(* IEC 61131-3 sources: plc-st-coding-agent/progress/evidence/f14_v3_parallel_20261112/jobs/custom_deepseek-v4pro (part 2) *)

(* ---- public-hard-05.raw_candidate_02.st ---- *)
FUNCTION_BLOCK MechanicalArmControl
VAR
    Step: INT := 1;                     // Current action step (1..8)
    ActionActive: BOOL := FALSE;        // TRUE when an automated action is being executed
    WaitingForStart: BOOL := TRUE;      // TRUE in single-step mode when waiting for start press
    CycleRunning: BOOL := FALSE;        // TRUE when a cycle is in progress (single/continuous)
    StartPrev: BOOL := FALSE;           // Previous value of Start input for edge detection
    StartPulse: BOOL := FALSE;          // One-scan pulse on rising edge of Start
    WaitingForStartPrev: BOOL := TRUE;  // Snapshot of WaitingForStart at scan start
    CycleRunningPrev: BOOL := FALSE;    // Snapshot of CycleRunning at scan start
END_VAR

// Rising edge detection for Start
StartPulse := Start AND NOT StartPrev;
StartPrev := Start;

// Capture previous states before any logic changes (to avoid race conditions)
WaitingForStartPrev := WaitingForStart;
CycleRunningPrev := CycleRunning;

IF NOT EmergencyStop THEN
    // Emergency stop triggered: stop all actions and reset automated state
    MoveDown := FALSE;
    MoveUp := FALSE;
    MoveLeft := FALSE;
    MoveRight := FALSE;
    ActivateGrip := FALSE;
    ActivateRelease := FALSE;
    Step := 1;
    ActionActive := FALSE;
    WaitingForStart := TRUE;
    CycleRunning := FALSE;
ELSE
    // Normal operation (no emergency stop)
    IF ManualMode THEN
        // Manual mode: direct button control with limit switch interlock
        MoveDown := DownButton AND NOT DownLimitSwitch;
        MoveUp := UpButton AND NOT UpLimitSwitch;
        MoveLeft := LeftButton AND NOT LeftLimitSwitch;
        MoveRight := RightButton AND NOT RightLimitSwitch;
        ActivateGrip := GripButton AND NOT GripLimitSwitch;
        ActivateRelease := ReleaseButton AND NOT ReleaseLimitSwitch;
        // Reset automated state when in manual mode
        Step := 1;
        ActionActive := FALSE;
        WaitingForStart := TRUE;
        CycleRunning := FALSE;
    ELSIF SingleStepMode THEN
        // Single step mode: one action per start press
        MoveDown := FALSE;
        MoveUp := FALSE;
        MoveLeft := FALSE;
        MoveRight := FALSE;
        ActivateGrip := FALSE;
        ActivateRelease := FALSE;

        IF WaitingForStartPrev AND StartPulse THEN
            WaitingForStart := FALSE;
            ActionActive := TRUE;
            Step := 1;  // Always start from step 1
        END_IF;

        IF ActionActive THEN
            CASE Step OF
                1: IF DownLimitSwitch THEN
                       ActionActive := FALSE;
                       WaitingForStart := TRUE;
                       Step := 1;
                   END_IF;
                2: IF GripLimitSwitch THEN
                       ActionActive := FALSE;
                       WaitingForStart := TRUE;
                       Step := 2;
                   END_IF;
                3: IF UpLimitSwitch THEN
                       ActionActive := FALSE;
                       WaitingForStart := TRUE;
                       Step := 3;
                   END_IF;
                4: IF RightLimitSwitch THEN
                       ActionActive := FALSE;
                       WaitingForStart := TRUE;
                       Step := 4;
                   END_IF;
                5: IF DownLimitSwitch THEN
                       ActionActive := FALSE;
                       WaitingForStart := TRUE;
                       Step := 5;
                   END_IF;
                6: IF ReleaseLimitSwitch THEN
                       ActionActive := FALSE;
                       WaitingForStart := TRUE;
                       Step := 6;
                   END_IF;
                7: IF UpLimitSwitch THEN
                       ActionActive := FALSE;
                       WaitingForStart := TRUE;
                       Step := 7;
                   END_IF;
                8: IF LeftLimitSwitch THEN
                       ActionActive := FALSE;
                       WaitingForStart := TRUE;
                       Step := 1;  // Reset to step 1 for next cycle
                   END_IF;
            END_CASE;
        END_IF;

        IF ActionActive THEN
            CASE Step OF
                1: MoveDown := TRUE;
                2: ActivateGrip := TRUE;
                3: MoveUp := TRUE;
                4: MoveRight := TRUE;
                5: MoveDown := TRUE;
                6: ActivateRelease := TRUE;
                7: MoveUp := TRUE;
                8: MoveLeft := TRUE;
            END_CASE;
        END_IF;
    ELSIF SingleCycleMode THEN
        // Single cycle mode: complete one full cycle automatically
        MoveDown := FALSE;
        MoveUp := FALSE;
        MoveLeft := FALSE;
        MoveRight := FALSE;
        ActivateGrip := FALSE;
        ActivateRelease := FALSE;

        IF NOT CycleRunningPrev AND StartPulse THEN
            CycleRunning := TRUE;
            Step := 1;
            ActionActive := TRUE;
        END_IF;

        IF CycleRunning AND ActionActive THEN
            CASE Step OF
                1: IF DownLimitSwitch THEN Step := 2; END_IF;
                2: IF GripLimitSwitch THEN Step := 3; END_IF;
                3: IF UpLimitSwitch THEN Step := 4; END_IF;
                4: IF RightLimitSwitch THEN Step := 5; END_IF;
                5: IF DownLimitSwitch THEN Step := 6; END_IF;
                6: IF ReleaseLimitSwitch THEN Step := 7; END_IF;
                7: IF UpLimitSwitch THEN Step := 8; END_IF;
                8: IF LeftLimitSwitch THEN
                       ActionActive := FALSE;   // Cycle finished
                       CycleRunning := FALSE;
                       Step := 1;               // Reset for next start
                   END_IF;
            END_CASE;
        END_IF;

        IF CycleRunning AND ActionActive THEN
            CASE Step OF
                1: MoveDown := TRUE;
                2: ActivateGrip := TRUE;
                3: MoveUp := TRUE;
                4: MoveRight := TRUE;
                5: MoveDown := TRUE;
                6: ActivateRelease := TRUE;
                7: MoveUp := TRUE;
                8: MoveLeft := TRUE;
            END_CASE;
        END_IF;
    ELSIF ContinuousMode THEN
        // Continuous mode: repeat cycle indefinitely
        MoveDown := FALSE;
        MoveUp := FALSE;
        MoveLeft := FALSE;
        MoveRight := FALSE;
        ActivateGrip := FALSE;
        ActivateRelease := FALSE;

        IF NOT CycleRunningPrev AND StartPulse THEN
            CycleRunning := TRUE;
            Step := 1;
            ActionActive := TRUE;
        END_IF;

        IF CycleRunning AND ActionActive THEN
            CASE Step OF
                1: IF DownLimitSwitch THEN Step := 2; END_IF;
                2: IF GripLimitSwitch THEN Step := 3; END_IF;
                3: IF UpLimitSwitch THEN Step := 4; END_IF;
                4: IF RightLimitSwitch THEN Step := 5; END_IF;
                5: IF DownLimitSwitch THEN Step := 6; END_IF;
                6: IF ReleaseLimitSwitch THEN Step := 7; END_IF;
                7: IF UpLimitSwitch THEN Step := 8; END_IF;
                8: IF LeftLimitSwitch THEN Step := 1; END_IF;  // Loop back
            END_CASE;
        END_IF;

        IF CycleRunning AND ActionActive THEN
            CASE Step OF
                1: MoveDown := TRUE;
                2: ActivateGrip := TRUE;
                3: MoveUp := TRUE;
                4: MoveRight := TRUE;
                5: MoveDown := TRUE;
                6: ActivateRelease := TRUE;
                7: MoveUp := TRUE;
                8: MoveLeft := TRUE;
            END_CASE;
        END_IF;
    ELSE
        // No mode selected (should not happen, but safe default)
        MoveDown := FALSE;
        MoveUp := FALSE;
        MoveLeft := FALSE;
        MoveRight := FALSE;
        ActivateGrip := FALSE;
        ActivateRelease := FALSE;
        Step := 1;
        ActionActive := FALSE;
        WaitingForStart := TRUE;
        CycleRunning := FALSE;
    END_IF;
END_IF;

END_FUNCTION_BLOCK

(* ---- public-hard-06.candidate_01.st ---- *)
TYPE T_PRODUCTION_STATE :
(
    IDLE,
    MOVING_FEED_TO_WASH,
    AT_WASH,
    MOVING_WASH_TO_WEIGHT,
    AT_WEIGHT_WAIT,
    AT_WEIGHT_REJECT,
    MOVING_WEIGHT_TO_FIRING,
    AT_FIRING,
    MOVING_FIRING_TO_OUTPUT,
    AT_OUTPUT
);
END_TYPE;

FUNCTION_BLOCK ProductionControl
VAR_INPUT
    Mode : BOOL;
    ForwardButton : BOOL;
    ReverseButton : BOOL;
    SensorFeed : BOOL;
    SensorWash : BOOL;
    SensorWeight : BOOL;
    SensorFiring : BOOL;
    SensorOutput : BOOL;
    washComplete : BOOL;
    weightComplete : BOOL;
    weight : REAL;
    firingComplete : BOOL;
END_VAR
VAR_OUTPUT
    MotorForward : BOOL;
    MotorReverse : BOOL;
    kick : BOOL;
    CompletionLight : BOOL;
    firingTemp : REAL;
END_VAR
VAR
    currentState : T_PRODUCTION_STATE := IDLE;
END_VAR

(* ---- public-hard-06.candidate_02.st ---- *)
TYPE T_PRODUCTION_STATE :
(
    IDLE,
    MOVING_FEED_TO_WASH,
    AT_WASH,
    MOVING_WASH_TO_WEIGHT,
    AT_WEIGHT_WAIT,
    AT_WEIGHT_REJECT,
    MOVING_WEIGHT_TO_FIRING,
    AT_FIRING,
    MOVING_FIRING_TO_OUTPUT,
    AT_OUTPUT
);
END_TYPE;

FUNCTION_BLOCK ProductionControl
VAR_INPUT
    Mode : BOOL;
    ForwardButton : BOOL;
    ReverseButton : BOOL;
    SensorFeed : BOOL;
    SensorWash : BOOL;
    SensorWeight : BOOL;
    SensorFiring : BOOL;
    SensorOutput : BOOL;
    washComplete : BOOL;
    weightComplete : BOOL;
    weight : REAL;
    firingComplete : BOOL;
END_VAR
VAR_OUTPUT
    MotorForward : BOOL;
    MotorReverse : BOOL;
    kick : BOOL;
    CompletionLight : BOOL;
    firingTemp : REAL;
END_VAR
VAR
    currentState : T_PRODUCTION_STATE := IDLE;
END_VAR

IF Mode = FALSE THEN
    // Manual mode
    IF ForwardButton AND NOT ReverseButton THEN
        MotorForward := TRUE;
        MotorReverse := FALSE;
    ELSIF ReverseButton AND NOT ForwardButton THEN
        MotorForward := FALSE;
        MotorReverse := TRUE;
    ELSE
        MotorForward := FALSE;
        MotorReverse := FALSE;
    END_IF;
    // Reset all automatic outputs and state
    kick := FALSE;
    CompletionLight := FALSE;
    firingTemp := 0.0;
    currentState := IDLE;
ELSE
    // Automatic mode
    // Set default outputs for this scan
    MotorReverse := FALSE;
    MotorForward := FALSE;
    kick := FALSE;
    CompletionLight := FALSE;
    // firingTemp retains its last calculated value unless updated in qualified weighing

    CASE currentState OF
        IDLE:
            IF SensorFeed THEN
                currentState := MOVING_FEED_TO_WASH;
                MotorForward := TRUE;
            END_IF;

        MOVING_FEED_TO_WASH:
            MotorForward := TRUE;
            IF SensorWash THEN
                MotorForward := FALSE;
                currentState := AT_WASH;
            END_IF;

        AT_WASH:
            IF washComplete THEN
                MotorForward := TRUE;
                currentState := MOVING_WASH_TO_WEIGHT;
            END_IF;

        MOVING_WASH_TO_WEIGHT:
            MotorForward := TRUE;
            IF SensorWeight THEN
                MotorForward := FALSE;
                currentState := AT_WEIGHT_WAIT;
            END_IF;

        AT_WEIGHT_WAIT:
            IF weightComplete THEN
                IF (weight >= 100.0) AND (weight <= 200.0) THEN
                    // Qualified material
                    firingTemp := 500.0 + (weight - 100.0) * 0.5;
                    MotorForward := TRUE;
                    currentState := MOVING_WEIGHT_TO_FIRING;
                ELSE
                    // Unqualified material
                    kick := TRUE;
                    currentState := AT_WEIGHT_REJECT;
                END_IF;
            END_IF;

        AT_WEIGHT_REJECT:
            kick := TRUE;
            IF NOT SensorWeight THEN
                kick := FALSE;
                currentState := IDLE;
            END_IF;

        MOVING_WEIGHT_TO_FIRING:
            MotorForward := TRUE;
            IF SensorFiring THEN
                MotorForward := FALSE;
                currentState := AT_FIRING;
            END_IF;

        AT_FIRING:
            IF firingComplete THEN
                MotorForward := TRUE;
                currentState := MOVING_FIRING_TO_OUTPUT;
            END_IF;

        MOVING_FIRING_TO_OUTPUT:
            MotorForward := TRUE;
            IF SensorOutput THEN
                MotorForward := FALSE;
                currentState := AT_OUTPUT;
            END_IF;

        AT_OUTPUT:
            CompletionLight := TRUE;
            IF NOT SensorOutput THEN
                CompletionLight := FALSE;
                currentState := IDLE;
            END_IF;
    END_CASE;
END_IF;

END_FUNCTION_BLOCK

(* ---- public-hard-06.raw_candidate_01.st ---- *)
TYPE T_PRODUCTION_STATE :
(
    IDLE,
    MOVING_FEED_TO_WASH,
    AT_WASH,
    MOVING_WASH_TO_WEIGHT,
    AT_WEIGHT_WAIT,
    AT_WEIGHT_REJECT,
    MOVING_WEIGHT_TO_FIRING,
    AT_FIRING,
    MOVING_FIRING_TO_OUTPUT,
    AT_OUTPUT
);
END_TYPE

FUNCTION_BLOCK ProductionControl
VAR_INPUT
    Mode : BOOL;
    ForwardButton : BOOL;
    ReverseButton : BOOL;
    SensorFeed : BOOL;
    SensorWash : BOOL;
    SensorWeight : BOOL;
    SensorFiring : BOOL;
    SensorOutput : BOOL;
    washComplete : BOOL;
    weightComplete : BOOL;
    weight : REAL;
    firingComplete : BOOL;
END_VAR
VAR_OUTPUT
    MotorForward : BOOL;
    MotorReverse : BOOL;
    kick : BOOL;
    CompletionLight : BOOL;
    firingTemp : REAL;
END_VAR
VAR
    currentState : T_PRODUCTION_STATE := IDLE;
END_VAR

(* ---- public-hard-06.raw_candidate_02.st ---- *)
TYPE T_PRODUCTION_STATE :
(
    IDLE,
    MOVING_FEED_TO_WASH,
    AT_WASH,
    MOVING_WASH_TO_WEIGHT,
    AT_WEIGHT_WAIT,
    AT_WEIGHT_REJECT,
    MOVING_WEIGHT_TO_FIRING,
    AT_FIRING,
    MOVING_FIRING_TO_OUTPUT,
    AT_OUTPUT
);
END_TYPE;

FUNCTION_BLOCK ProductionControl
VAR_INPUT
    Mode : BOOL;
    ForwardButton : BOOL;
    ReverseButton : BOOL;
    SensorFeed : BOOL;
    SensorWash : BOOL;
    SensorWeight : BOOL;
    SensorFiring : BOOL;
    SensorOutput : BOOL;
    washComplete : BOOL;
    weightComplete : BOOL;
    weight : REAL;
    firingComplete : BOOL;
END_VAR
VAR_OUTPUT
    MotorForward : BOOL;
    MotorReverse : BOOL;
    kick : BOOL;
    CompletionLight : BOOL;
    firingTemp : REAL;
END_VAR
VAR
    currentState : T_PRODUCTION_STATE := IDLE;
END_VAR

IF Mode = FALSE THEN
    // Manual mode
    IF ForwardButton AND NOT ReverseButton THEN
        MotorForward := TRUE;
        MotorReverse := FALSE;
    ELSIF ReverseButton AND NOT ForwardButton THEN
        MotorForward := FALSE;
        MotorReverse := TRUE;
    ELSE
        MotorForward := FALSE;
        MotorReverse := FALSE;
    END_IF;
    // Reset all automatic outputs and state
    kick := FALSE;
    CompletionLight := FALSE;
    firingTemp := 0.0;
    currentState := IDLE;
ELSE
    // Automatic mode
    // Set default outputs for this scan
    MotorReverse := FALSE;
    MotorForward := FALSE;
    kick := FALSE;
    CompletionLight := FALSE;
    // firingTemp retains its last calculated value unless updated in qualified weighing

    CASE currentState OF
        IDLE:
            IF SensorFeed THEN
                currentState := MOVING_FEED_TO_WASH;
                MotorForward := TRUE;
            END_IF;

        MOVING_FEED_TO_WASH:
            MotorForward := TRUE;
            IF SensorWash THEN
                MotorForward := FALSE;
                currentState := AT_WASH;
            END_IF;

        AT_WASH:
            IF washComplete THEN
                MotorForward := TRUE;
                currentState := MOVING_WASH_TO_WEIGHT;
            END_IF;

        MOVING_WASH_TO_WEIGHT:
            MotorForward := TRUE;
            IF SensorWeight THEN
                MotorForward := FALSE;
                currentState := AT_WEIGHT_WAIT;
            END_IF;

        AT_WEIGHT_WAIT:
            IF weightComplete THEN
                IF (weight >= 100.0) AND (weight <= 200.0) THEN
                    // Qualified material
                    firingTemp := 500.0 + (weight - 100.0) * 0.5;
                    MotorForward := TRUE;
                    currentState := MOVING_WEIGHT_TO_FIRING;
                ELSE
                    // Unqualified material
                    kick := TRUE;
                    currentState := AT_WEIGHT_REJECT;
                END_IF;
            END_IF;

        AT_WEIGHT_REJECT:
            kick := TRUE;
            IF NOT SensorWeight THEN
                kick := FALSE;
                currentState := IDLE;
            END_IF;

        MOVING_WEIGHT_TO_FIRING:
            MotorForward := TRUE;
            IF SensorFiring THEN
                MotorForward := FALSE;
                currentState := AT_FIRING;
            END_IF;

        AT_FIRING:
            IF firingComplete THEN
                MotorForward := TRUE;
                currentState := MOVING_FIRING_TO_OUTPUT;
            END_IF;

        MOVING_FIRING_TO_OUTPUT:
            MotorForward := TRUE;
            IF SensorOutput THEN
                MotorForward := FALSE;
                currentState := AT_OUTPUT;
            END_IF;

        AT_OUTPUT:
            CompletionLight := TRUE;
            IF NOT SensorOutput THEN
                CompletionLight := FALSE;
                currentState := IDLE;
            END_IF;
    END_CASE;
END_IF;

END_FUNCTION_BLOCK

(* ---- public-medium-01.candidate_01.st ---- *)
TYPE ST_Pump :
STRUCT
    priority : INT;
    selection : BOOL;
    RunComd : BOOL;
END_STRUCT;
END_TYPE;

FUNCTION_BLOCK FB_MultiPumpControl
VAR_INPUT
    mode : BOOL;
    start : BOOL;
    stop : BOOL;
END_VAR
VAR_IN_OUT
    pumpGroup : ARRAY[1..5] OF ST_Pump;
END_VAR
VAR
    runActive : BOOL := FALSE;
    autoSelected : ARRAY[1..5] OF BOOL;
    i : INT;
    j : INT;
    rank : INT;
END_VAR

IF stop THEN
    runActive := FALSE;
    FOR i := 1 TO 5 DO
        pumpGroup[i].RunComd := FALSE;
    END_FOR;
ELSE
    IF start THEN
        runActive := TRUE;
    END_IF;

    IF runActive THEN
        IF mode THEN
            FOR i := 1 TO 5 DO
                rank := 0;
                FOR j := 1 TO 5 DO
                    IF (pumpGroup[j].priority > pumpGroup[i].priority) OR
                       ((pumpGroup[j].priority = pumpGroup[i].priority) AND (j < i)) THEN
                        rank := rank + 1;
                    END_IF;
                END_FOR;
                autoSelected[i] := (rank < 3);
            END_FOR;

            FOR i := 1 TO 5 DO
                pumpGroup[i].RunComd := autoSelected[i];
            END_FOR;
        ELSE
            FOR i := 1 TO 5 DO
                pumpGroup[i].RunComd := pumpGroup[i].selection;
            END_FOR;
        END_IF;
    ELSE
        FOR i := 1 TO 5 DO
            pumpGroup[i].RunComd := FALSE;
        END_FOR;
    END_IF;
END_IF;

END_FUNCTION_BLOCK

(* ---- public-medium-01.candidate_02.st ---- *)
TYPE ST_Pump :
STRUCT
    priority : INT;
    selection : BOOL;
    RunComd : BOOL;
END_STRUCT;
END_TYPE;

FUNCTION_BLOCK FB_MultiPumpControl
VAR_INPUT
    mode : BOOL;
    start : BOOL;
    stop : BOOL;
END_VAR
VAR_IN_OUT
    pumpGroup : ARRAY[1..5] OF ST_Pump;
END_VAR
VAR
    runActive : BOOL := FALSE;
    autoSelected : ARRAY[1..5] OF BOOL;
    i : INT;
    j : INT;
    rank : INT;
END_VAR

IF stop THEN
    runActive := FALSE;
    FOR i := 1 TO 5 DO
        pumpGroup[i].RunComd := FALSE;
    END_FOR;
ELSE
    IF start THEN
        runActive := TRUE;
    END_IF;

    IF runActive THEN
        IF mode THEN
            FOR i := 1 TO 5 DO
                rank := 0;
                FOR j := 1 TO 5 DO
                    IF (pumpGroup[j].priority > pumpGroup[i].priority) OR
                       ((pumpGroup[j].priority = pumpGroup[i].priority) AND (j < i)) THEN
                        rank := rank + 1;
                    END_IF;
                END_FOR;
                autoSelected[i] := (rank < 3);
            END_FOR;

            FOR i := 1 TO 5 DO
                pumpGroup[i].RunComd := autoSelected[i];
            END_FOR;
        ELSE
            FOR i := 1 TO 5 DO
                pumpGroup[i].RunComd := pumpGroup[i].selection;
            END_FOR;
        END_IF;
    ELSE
        FOR i := 1 TO 5 DO
            pumpGroup[i].RunComd := FALSE;
        END_FOR;
    END_IF;
END_IF;

END_FUNCTION_BLOCK

(* ---- public-medium-01.raw_candidate_01.st ---- *)
TYPE ST_Pump :
STRUCT
    priority : INT;
    selection : BOOL;
    RunComd : BOOL;
END_STRUCT;
END_TYPE;

FUNCTION_BLOCK FB_MultiPumpControl
VAR_INPUT
    mode : BOOL;
    start : BOOL;
    stop : BOOL;
END_VAR
VAR_IN_OUT
    pumpGroup : ARRAY[1..5] OF ST_Pump;
END_VAR
VAR
    runActive : BOOL := FALSE;
    autoSelected : ARRAY[1..5] OF BOOL;
    i : INT;
    j : INT;
    rank : INT;
END_VAR

IF stop THEN
    runActive := FALSE;
    FOR i := 1 TO 5 DO
        pumpGroup[i].RunComd := FALSE;
    END_FOR;
ELSE
    IF start THEN
        runActive := TRUE;
    END_IF;

    IF runActive THEN
        IF mode THEN
            FOR i := 1 TO 5 DO
                rank := 0;
                FOR j := 1 TO 5 DO
                    IF (pumpGroup[j].priority > pumpGroup[i].priority) OR
                       ((pumpGroup[j].priority = pumpGroup[i].priority) AND (j < i)) THEN
                        rank := rank + 1;
                    END_IF;
                END_FOR;
                autoSelected[i] := (rank < 3);
            END_FOR;

            FOR i := 1 TO 5 DO
                pumpGroup[i].RunComd := autoSelected[i];
            END_FOR;
        ELSE
            FOR i := 1 TO 5 DO
                pumpGroup[i].RunComd := pumpGroup[i].selection;
            END_FOR;
        END_IF;
    ELSE
        FOR i := 1 TO 5 DO
            pumpGroup[i].RunComd := FALSE;
        END_FOR;
    END_IF;
END_IF;

END_FUNCTION_BLOCK

(* ---- public-medium-01.raw_candidate_02.st ---- *)
TYPE ST_Pump :
STRUCT
    priority : INT;
    selection : BOOL;
    RunComd : BOOL;
END_STRUCT
END_TYPE

FUNCTION_BLOCK FB_MultiPumpControl
VAR_INPUT
    mode : BOOL;
    start : BOOL;
    stop : BOOL;
END_VAR
VAR_IN_OUT
    pumpGroup : ARRAY[1..5] OF ST_Pump;
END_VAR
VAR
    runActive : BOOL := FALSE;
    autoSelected : ARRAY[1..5] OF BOOL;
    i : INT;
    j : INT;
    rank : INT;
END_VAR

IF stop THEN
    runActive := FALSE;
    FOR i := 1 TO 5 DO
        pumpGroup[i].RunComd := FALSE;
    END_FOR;
ELSE
    IF start THEN
        runActive := TRUE;
    END_IF;

    IF runActive THEN
        IF mode THEN
            FOR i := 1 TO 5 DO
                rank := 0;
                FOR j := 1 TO 5 DO
                    IF (pumpGroup[j].priority > pumpGroup[i].priority) OR
                       ((pumpGroup[j].priority = pumpGroup[i].priority) AND (j < i)) THEN
                        rank := rank + 1;
                    END_IF;
                END_FOR;
                autoSelected[i] := (rank < 3);
            END_FOR;

            FOR i := 1 TO 5 DO
                pumpGroup[i].RunComd := autoSelected[i];
            END_FOR;
        ELSE
            FOR i := 1 TO 5 DO
                pumpGroup[i].RunComd := pumpGroup[i].selection;
            END_FOR;
        END_IF;
    ELSE
        FOR i := 1 TO 5 DO
            pumpGroup[i].RunComd := FALSE;
        END_FOR;
    END_IF;
END_IF;

END_FUNCTION_BLOCK

(* ---- public-medium-02.candidate_01.st ---- *)
TYPE ST_AnalogChannel :
STRUCT
    enable : BOOL;
    hiLIM : REAL;
    loLIM : REAL;
    bipolar : BOOL;
    measuringMode : INT;
    retVal : WORD;
    outputValue : REAL;
END_STRUCT;
END_TYPE;

FUNCTION_BLOCK AnalogBatchProcessing
VAR_INPUT
    count : DINT;
END_VAR
VAR_INOUT
    analogValues : ARRAY[*] OF INT;
    channels : ARRAY[*] OF ST_AnalogChannel;
END_VAR
VAR
    i : DINT;
    idxA : DINT;
    idxC : DINT;
    lbA : DINT;
    lbC : DINT;
    raw : INT;
    rawReal : REAL;
    rawMin : REAL;
    rawSpan : REAL;
    engSpan : REAL;
END_VAR

    lbA := LOWER_BOUND(analogValues, 1);
    lbC := LOWER_BOUND(channels, 1);

    FOR i := 0 TO count - 1 DO
        idxA := lbA + i;
        idxC := lbC + i;
        raw := analogValues[idxA];
        channels[idxC].retVal := 0;

        IF channels[idxC].enable THEN
            IF channels[idxC].measuringMode <> 0 AND channels[idxC].measuringMode <> 1 AND channels[idxC].measuringMode <> 2 THEN
                channels[idxC].retVal := WORD#16#8001;
            ELSIF channels[idxC].hiLIM <= channels[idxC].loLIM THEN
                channels[idxC].retVal := WORD#16#8002;
            ELSIF channels[idxC].measuringMode = 0 THEN
                rawReal := INT_TO_REAL(raw);

                IF channels[idxC].bipolar THEN
                    rawMin := -27648.0;
                    rawSpan := 55296.0;
                ELSE
                    rawMin := 0.0;
                    rawSpan := 27648.0;
                END_IF;

                engSpan := channels[idxC].hiLIM - channels[idxC].loLIM;
                channels[idxC].outputValue := channels[idxC].loLIM + (rawReal - rawMin) * engSpan / rawSpan;
            ELSIF channels[idxC].measuringMode = 1 THEN
                rawReal := INT_TO_REAL(raw);
                channels[idxC].outputValue := rawReal / 10.0;
            ELSE
                rawReal := INT_TO_REAL(raw);
                channels[idxC].outputValue := rawReal / 100.0;
            END_IF;
        END_IF;
    END_FOR;

END_FUNCTION_BLOCK

(* ---- public-medium-02.candidate_02.st ---- *)
TYPE ST_AnalogChannel :
STRUCT
    enable : BOOL;
    hiLIM : REAL;
    loLIM : REAL;
    bipolar : BOOL;
    measuringMode : INT;
    retVal : WORD;
    outputValue : REAL;
END_STRUCT;
END_TYPE;

FUNCTION_BLOCK AnalogBatchProcessing
VAR_INPUT
    count : DINT;
END_VAR
VAR_IN_OUT
    analogValues : ARRAY[*] OF INT;
    channels : ARRAY[*] OF ST_AnalogChannel;
END_VAR
VAR
    i : DINT;
    idxA : DINT;
    idxC : DINT;
    lbA : DINT;
    lbC : DINT;
    raw : INT;
    rawReal : REAL;
    rawMin : REAL;
    rawSpan : REAL;
    engSpan : REAL;
END_VAR

    lbA := LOWER_BOUND(analogValues, 1);
    lbC := LOWER_BOUND(channels, 1);

    FOR i := 0 TO count - 1 DO
        idxA := lbA + i;
        idxC := lbC + i;

        IF channels[idxC].enable THEN
            IF channels[idxC].measuringMode <> 0 AND channels[idxC].measuringMode <> 1 AND channels[idxC].measuringMode <> 2 THEN
                channels[idxC].retVal := WORD#16#8001;
            ELSIF channels[idxC].hiLIM <= channels[idxC].loLIM THEN
                channels[idxC].retVal := WORD#16#8002;
            ELSE
                raw := analogValues[idxA];
                rawReal := INT_TO_REAL(raw);
                CASE channels[idxC].measuringMode OF
                    0:
                        IF channels[idxC].bipolar THEN
                            rawMin := -27648.0;
                            rawSpan := 55296.0;
                        ELSE
                            rawMin := 0.0;
                            rawSpan := 27648.0;
                        END_IF;
                        engSpan := channels[idxC].hiLIM - channels[idxC].loLIM;
                        channels[idxC].outputValue := channels[idxC].loLIM + (rawReal - rawMin) * engSpan / rawSpan;
                    1:
                        channels[idxC].outputValue := rawReal / 10.0;
                    2:
                        channels[idxC].outputValue := rawReal / 100.0;
                END_CASE;
                channels[idxC].retVal := 0;
            END_IF;
        END_IF;
    END_FOR;

END_FUNCTION_BLOCK

(* ---- public-medium-02.raw_candidate_01.st ---- *)
TYPE ST_AnalogChannel :
STRUCT
    enable : BOOL;
    hiLIM : REAL;
    loLIM : REAL;
    bipolar : BOOL;
    measuringMode : INT;
    retVal : WORD;
    outputValue : REAL;
END_STRUCT
END_TYPE

FUNCTION_BLOCK AnalogBatchProcessing
VAR_INPUT
    count : DINT;
END_VAR
VAR_INOUT
    analogValues : ARRAY[*] OF INT;
    channels : ARRAY[*] OF ST_AnalogChannel;
END_VAR
VAR
    i : DINT;
    idxA : DINT;
    idxC : DINT;
    lbA : DINT;
    lbC : DINT;
    raw : INT;
    rawReal : REAL;
    rawMin : REAL;
    rawSpan : REAL;
    engSpan : REAL;
END_VAR

    lbA := LOWER_BOUND(analogValues, 1);
    lbC := LOWER_BOUND(channels, 1);

    FOR i := 0 TO count - 1 DO
        idxA := lbA + i;
        idxC := lbC + i;
        raw := analogValues[idxA];
        channels[idxC].retVal := 0;

        IF channels[idxC].enable THEN
            IF channels[idxC].measuringMode <> 0 AND channels[idxC].measuringMode <> 1 AND channels[idxC].measuringMode <> 2 THEN
                channels[idxC].retVal := WORD#16#8001;
            ELSIF channels[idxC].hiLIM <= channels[idxC].loLIM THEN
                channels[idxC].retVal := WORD#16#8002;
            ELSIF channels[idxC].measuringMode = 0 THEN
                rawReal := INT_TO_REAL(raw);

                IF channels[idxC].bipolar THEN
                    rawMin := -27648.0;
                    rawSpan := 55296.0;
                ELSE
                    rawMin := 0.0;
                    rawSpan := 27648.0;
                END_IF

                engSpan := channels[idxC].hiLIM - channels[idxC].loLIM;
                channels[idxC].outputValue := channels[idxC].loLIM + (rawReal - rawMin) * engSpan / rawSpan;
            ELSIF channels[idxC].measuringMode = 1 THEN
                rawReal := INT_TO_REAL(raw);
                channels[idxC].outputValue := rawReal / 10.0;
            ELSE
                rawReal := INT_TO_REAL(raw);
                channels[idxC].outputValue := rawReal / 100.0;
            END_IF
        END_IF
    END_FOR

END_FUNCTION_BLOCK

(* ---- public-medium-02.raw_candidate_02.st ---- *)
TYPE ST_AnalogChannel :
STRUCT
    enable : BOOL;
    hiLIM : REAL;
    loLIM : REAL;
    bipolar : BOOL;
    measuringMode : INT;
    retVal : WORD;
    outputValue : REAL;
END_STRUCT;
END_TYPE;

FUNCTION_BLOCK AnalogBatchProcessing
VAR_INPUT
    count : DINT;
END_VAR
VAR_IN_OUT
    analogValues : ARRAY[*] OF INT;
    channels : ARRAY[*] OF ST_AnalogChannel;
END_VAR
VAR
    i : DINT;
    idxA : DINT;
    idxC : DINT;
    lbA : DINT;
    lbC : DINT;
    raw : INT;
    rawReal : REAL;
    rawMin : REAL;
    rawSpan : REAL;
    engSpan : REAL;
END_VAR

    lbA := LOWER_BOUND(analogValues, 1);
    lbC := LOWER_BOUND(channels, 1);

    FOR i := 0 TO count - 1 DO
        idxA := lbA + i;
        idxC := lbC + i;

        IF channels[idxC].enable THEN
            IF channels[idxC].measuringMode <> 0 AND channels[idxC].measuringMode <> 1 AND channels[idxC].measuringMode <> 2 THEN
                channels[idxC].retVal := WORD#16#8001;
            ELSIF channels[idxC].hiLIM <= channels[idxC].loLIM THEN
                channels[idxC].retVal := WORD#16#8002;
            ELSE
                raw := analogValues[idxA];
                rawReal := INT_TO_REAL(raw);
                CASE channels[idxC].measuringMode OF
                    0:
                        IF channels[idxC].bipolar THEN
                            rawMin := -27648.0;
                            rawSpan := 55296.0;
                        ELSE
                            rawMin := 0.0;
                            rawSpan := 27648.0;
                        END_IF;
                        engSpan := channels[idxC].hiLIM - channels[idxC].loLIM;
                        channels[idxC].outputValue := channels[idxC].loLIM + (rawReal - rawMin) * engSpan / rawSpan;
                    1:
                        channels[idxC].outputValue := rawReal / 10.0;
                    2:
                        channels[idxC].outputValue := rawReal / 100.0;
                END_CASE;
                channels[idxC].retVal := 0;
            END_IF;
        END_IF;
    END_FOR;

END_FUNCTION_BLOCK

(* ---- public-medium-03.candidate_01.st ---- *)
FUNCTION_BLOCK FB_MovingAverage
VAR_INPUT
    cyclicExecution : BOOL;
    trigger : BOOL;
    value : LREAL;
    windowSize : INT;
    reset : BOOL;
END_VAR
VAR_OUTPUT
    average : LREAL;
    windowSizeReached : BOOL;
    error : BOOL;
    status : WORD;
END_VAR
VAR
    buffer : ARRAY[0..99] OF LREAL;
    count : INT := 0;
    writeIndex : INT := 0;
    sum : LREAL := 0.0;
    prevTrigger : BOOL := FALSE;
    prevWindowSize : INT := 0;
    updateNow : BOOL;
END_VAR

IF (windowSize < 1) OR (windowSize > 100) THEN
    error := TRUE;
    status := 16#8200;
    average := 0.0;
    windowSizeReached := FALSE;
    count := 0;
    writeIndex := 0;
    sum := 0.0;
ELSE
    error := FALSE;
    status := 16#0000;

    IF reset OR (windowSize <> prevWindowSize) THEN
        count := 0;
        writeIndex := 0;
        sum := 0.0;
        average := 0.0;
        windowSizeReached := FALSE;
    END_IF;
    prevWindowSize := windowSize;

    IF cyclicExecution THEN
        updateNow := TRUE;
    ELSIF (trigger AND NOT prevTrigger) THEN
        updateNow := TRUE;
    ELSE
        updateNow := FALSE;
    END_IF;

    IF updateNow THEN
        IF count < windowSize THEN
            buffer[writeIndex] := value;
            sum := sum + value;
            count := count + 1;
            writeIndex := writeIndex + 1;
        ELSE
            sum := sum - buffer[writeIndex] + value;
            buffer[writeIndex] := value;
            writeIndex := (writeIndex + 1) MOD windowSize;
        END_IF;
        IF count > 0 THEN
            average := sum / count;
        ELSE
            average := 0.0;
        END_IF;
        windowSizeReached := (count >= windowSize);
    END_IF;
END_IF;

prevTrigger := trigger;

(* ---- public-medium-03.candidate_02.st ---- *)
FUNCTION_BLOCK FB_MovingAverage
VAR_INPUT
    cyclicExecution : BOOL;
    trigger : BOOL;
    value : LREAL;
    windowSize : INT;
    reset : BOOL;
END_VAR
VAR_OUTPUT
    average : LREAL;
    windowSizeReached : BOOL;
    error : BOOL;
    status : WORD;
END_VAR
VAR
    buffer : ARRAY[0..99] OF LREAL;
    count : INT := 0;
    writeIndex : INT := 0;
    sum : LREAL := 0.0;
    prevTrigger : BOOL := FALSE;
    prevWindowSize : INT := 0;
    updateNow : BOOL;
END_VAR

IF (windowSize < 1) OR (windowSize > 100) THEN
    error := TRUE;
    status := 16#8200;
    average := 0.0;
    windowSizeReached := FALSE;
    count := 0;
    writeIndex := 0;
    sum := 0.0;
ELSE
    error := FALSE;
    status := 16#0000;

    IF reset OR (windowSize <> prevWindowSize) THEN
        count := 0;
        writeIndex := 0;
        sum := 0.0;
        average := 0.0;
        windowSizeReached := FALSE;
    END_IF;
    prevWindowSize := windowSize;

    IF cyclicExecution THEN
        updateNow := TRUE;
    ELSIF (trigger AND NOT prevTrigger) THEN
        updateNow := TRUE;
    ELSE
        updateNow := FALSE;
    END_IF;

    IF updateNow THEN
        IF count < windowSize THEN
            buffer[writeIndex] := value;
            sum := sum + value;
            count := count + 1;
            writeIndex := (writeIndex + 1) MOD windowSize;
        ELSE
            sum := sum - buffer[writeIndex] + value;
            buffer[writeIndex] := value;
            writeIndex := (writeIndex + 1) MOD windowSize;
        END_IF;
        IF count > 0 THEN
            average := sum / count;
        ELSE
            average := 0.0;
        END_IF;
        windowSizeReached := (count >= windowSize);
    END_IF;
END_IF;

prevTrigger := trigger;

END_FUNCTION_BLOCK

(* ---- public-medium-03.raw_candidate_01.st ---- *)
FUNCTION_BLOCK FB_MovingAverage
VAR_INPUT
    cyclicExecution : BOOL;
    trigger : BOOL;
    value : LREAL;
    windowSize : INT;
    reset : BOOL;
END_VAR
VAR_OUTPUT
    average : LREAL;
    windowSizeReached : BOOL;
    error : BOOL;
    status : WORD;
END_VAR
VAR
    buffer : ARRAY[0..99] OF LREAL;
    count : INT := 0;
    writeIndex : INT := 0;
    sum : LREAL := 0.0;
    prevTrigger : BOOL := FALSE;
    prevWindowSize : INT := 0;
    updateNow : BOOL;
END_VAR

IF (windowSize < 1) OR (windowSize > 100) THEN
    error := TRUE;
    status := 16#8200;
    average := 0.0;
    windowSizeReached := FALSE;
    count := 0;
    writeIndex := 0;
    sum := 0.0;
ELSE
    error := FALSE;
    status := 16#0000;

    IF reset OR (windowSize <> prevWindowSize) THEN
        count := 0;
        writeIndex := 0;
        sum := 0.0;
        average := 0.0;
        windowSizeReached := FALSE;
    END_IF;
    prevWindowSize := windowSize;

    IF cyclicExecution THEN
        updateNow := TRUE;
    ELSIF (trigger AND NOT prevTrigger) THEN
        updateNow := TRUE;
    ELSE
        updateNow := FALSE;
    END_IF;

    IF updateNow THEN
        IF count < windowSize THEN
            buffer[writeIndex] := value;
            sum := sum + value;
            count := count + 1;
            writeIndex := writeIndex + 1;
        ELSE
            sum := sum - buffer[writeIndex] + value;
            buffer[writeIndex] := value;
            writeIndex := (writeIndex + 1) MOD windowSize;
        END_IF;
        IF count > 0 THEN
            average := sum / count;
        ELSE
            average := 0.0;
        END_IF;
        windowSizeReached := (count >= windowSize);
    END_IF;
END_IF;

prevTrigger := trigger;

(* ---- public-medium-03.raw_candidate_02.st ---- *)
FUNCTION_BLOCK FB_MovingAverage
VAR_INPUT
    cyclicExecution : BOOL;
    trigger : BOOL;
    value : LREAL;
    windowSize : INT;
    reset : BOOL;
END_VAR
VAR_OUTPUT
    average : LREAL;
    windowSizeReached : BOOL;
    error : BOOL;
    status : WORD;
END_VAR
VAR
    buffer : ARRAY[0..99] OF LREAL;
    count : INT := 0;
    writeIndex : INT := 0;
    sum : LREAL := 0.0;
    prevTrigger : BOOL := FALSE;
    prevWindowSize : INT := 0;
    updateNow : BOOL;
END_VAR

IF (windowSize < 1) OR (windowSize > 100) THEN
    error := TRUE;
    status := 16#8200;
    average := 0.0;
    windowSizeReached := FALSE;
    count := 0;
    writeIndex := 0;
    sum := 0.0;
ELSE
    error := FALSE;
    status := 16#0000;

    IF reset OR (windowSize <> prevWindowSize) THEN
        count := 0;
        writeIndex := 0;
        sum := 0.0;
        average := 0.0;
        windowSizeReached := FALSE;
    END_IF;
    prevWindowSize := windowSize;

    IF cyclicExecution THEN
        updateNow := TRUE;
    ELSIF (trigger AND NOT prevTrigger) THEN
        updateNow := TRUE;
    ELSE
        updateNow := FALSE;
    END_IF;

    IF updateNow THEN
        IF count < windowSize THEN
            buffer[writeIndex] := value;
            sum := sum + value;
            count := count + 1;
            writeIndex := (writeIndex + 1) MOD windowSize;
        ELSE
            sum := sum - buffer[writeIndex] + value;
            buffer[writeIndex] := value;
            writeIndex := (writeIndex + 1) MOD windowSize;
        END_IF;
        IF count > 0 THEN
            average := sum / count;
        ELSE
            average := 0.0;
        END_IF;
        windowSizeReached := (count >= windowSize);
    END_IF;
END_IF;

prevTrigger := trigger;

END_FUNCTION_BLOCK

(* ---- public-medium-04.candidate_01.st ---- *)
FUNCTION_BLOCK FB_TemperatureLogicControl
VAR_INPUT
    TemperatureSensorInput : REAL;
    SetTemperature : REAL;
END_VAR
VAR_OUTPUT
    CurrentTemperature : REAL;
    SetTempDisplay : REAL;
    HeaterStatus : BOOL;
    OverheatProtection : BOOL;
    HeaterOutput : BOOL;
END_VAR
VAR
    heaterOnTimer : TON;
    coolingTimer : TON;
    SensorFault : BOOL;
END_VAR

CurrentTemperature := TemperatureSensorInput;
SetTempDisplay := SetTemperature;

SensorFault := (TemperatureSensorInput < 0.0) OR (TemperatureSensorInput > 100.0);

heaterOnTimer(IN := HeaterOutput, PT := T#5S);

IF (NOT SensorFault) AND (NOT OverheatProtection) AND heaterOnTimer.Q THEN
    OverheatProtection := TRUE;
END_IF;

coolingTimer(IN := OverheatProtection, PT := T#3S);

IF OverheatProtection THEN
    HeaterOutput := FALSE;
    IF coolingTimer.Q THEN
        OverheatProtection := FALSE;
    END_IF;
ELSIF SensorFault THEN
    HeaterOutput := FALSE;
ELSIF TemperatureSensorInput < SetTemperature THEN
    HeaterOutput := TRUE;
ELSE
    HeaterOutput := FALSE;
END_IF;

HeaterStatus := HeaterOutput;

(* ---- public-medium-04.candidate_02.st ---- *)
FUNCTION_BLOCK FB_TemperatureLogicControl
VAR_INPUT
    TemperatureSensorInput : REAL;
    SetTemperature : REAL;
END_VAR
VAR_OUTPUT
    CurrentTemperature : REAL;
    SetTempDisplay : REAL;
    HeaterStatus : BOOL;
    OverheatProtection : BOOL;
    HeaterOutput : BOOL;
END_VAR
VAR
    heaterOnTimer : TON;
    coolingTimer : TON;
    SensorFault : BOOL;
END_VAR

CurrentTemperature := TemperatureSensorInput;
SetTempDisplay := SetTemperature;

SensorFault := (TemperatureSensorInput < 0.0) OR (TemperatureSensorInput > 100.0);

heaterOnTimer(IN := HeaterOutput, PT := T#5S);
IF (NOT SensorFault) AND (NOT OverheatProtection) AND heaterOnTimer.Q THEN
    OverheatProtection := TRUE;
END_IF;

coolingTimer(IN := OverheatProtection, PT := T#3S);

IF OverheatProtection THEN
    HeaterOutput := FALSE;
    IF coolingTimer.Q THEN
        OverheatProtection := FALSE;
    END_IF;
ELSIF SensorFault THEN
    HeaterOutput := FALSE;
ELSIF TemperatureSensorInput < SetTemperature THEN
    HeaterOutput := TRUE;
ELSE
    HeaterOutput := FALSE;
END_IF;

HeaterStatus := HeaterOutput;

END_FUNCTION_BLOCK

(* ---- public-medium-04.raw_candidate_01.st ---- *)
FUNCTION_BLOCK FB_TemperatureLogicControl
VAR_INPUT
    TemperatureSensorInput : REAL;
    SetTemperature : REAL;
END_VAR
VAR_OUTPUT
    CurrentTemperature : REAL;
    SetTempDisplay : REAL;
    HeaterStatus : BOOL;
    OverheatProtection : BOOL;
    HeaterOutput : BOOL;
END_VAR
VAR
    heaterOnTimer : TON;
    coolingTimer : TON;
    SensorFault : BOOL;
END_VAR

CurrentTemperature := TemperatureSensorInput;
SetTempDisplay := SetTemperature;

SensorFault := (TemperatureSensorInput < 0.0) OR (TemperatureSensorInput > 100.0);

heaterOnTimer(IN := HeaterOutput, PT := T#5S);

IF (NOT SensorFault) AND (NOT OverheatProtection) AND heaterOnTimer.Q THEN
    OverheatProtection := TRUE;
END_IF;

coolingTimer(IN := OverheatProtection, PT := T#3S);

IF OverheatProtection THEN
    HeaterOutput := FALSE;
    IF coolingTimer.Q THEN
        OverheatProtection := FALSE;
    END_IF;
ELSIF SensorFault THEN
    HeaterOutput := FALSE;
ELSIF TemperatureSensorInput < SetTemperature THEN
    HeaterOutput := TRUE;
ELSE
    HeaterOutput := FALSE;
END_IF;

HeaterStatus := HeaterOutput;

(* ---- public-medium-04.raw_candidate_02.st ---- *)
FUNCTION_BLOCK FB_TemperatureLogicControl
VAR_INPUT
    TemperatureSensorInput : REAL;
    SetTemperature : REAL;
END_VAR
VAR_OUTPUT
    CurrentTemperature : REAL;
    SetTempDisplay : REAL;
    HeaterStatus : BOOL;
    OverheatProtection : BOOL;
    HeaterOutput : BOOL;
END_VAR
VAR
    heaterOnTimer : TON;
    coolingTimer : TON;
    SensorFault : BOOL;
END_VAR

CurrentTemperature := TemperatureSensorInput;
SetTempDisplay := SetTemperature;

SensorFault := (TemperatureSensorInput < 0.0) OR (TemperatureSensorInput > 100.0);

heaterOnTimer(IN := HeaterOutput, PT := T#5S);
IF (NOT SensorFault) AND (NOT OverheatProtection) AND heaterOnTimer.Q THEN
    OverheatProtection := TRUE;
END_IF;

coolingTimer(IN := OverheatProtection, PT := T#3S);

IF OverheatProtection THEN
    HeaterOutput := FALSE;
    IF coolingTimer.Q THEN
        OverheatProtection := FALSE;
    END_IF;
ELSIF SensorFault THEN
    HeaterOutput := FALSE;
ELSIF TemperatureSensorInput < SetTemperature THEN
    HeaterOutput := TRUE;
ELSE
    HeaterOutput := FALSE;
END_IF;

HeaterStatus := HeaterOutput;

END_FUNCTION_BLOCK

(* ---- public-medium-05.candidate_01.st ---- *)
TYPE AutoState : (IDLE, MOVING_TO_B, WAIT_B, MOVING_TO_C, WAIT_C);
END_TYPE;

FUNCTION_BLOCK ProductionLineControl
VAR_INPUT
    Mode : BOOL;
    ForwardButton : BOOL;
    ReverseButton : BOOL;
    SensorA : BOOL;
    SensorB : BOOL;
    SensorC : BOOL;
    ButtonA : BOOL;
    ButtonB : BOOL;
    ButtonC : BOOL;
END_VAR
VAR_OUTPUT
    MotorForward : BOOL;
    MotorReverse : BOOL;
    CompletionLight : BOOL;
END_VAR
VAR
    State : AutoState := IDLE;
    CompletionLatched : BOOL := FALSE;
END_VAR

MotorForward := FALSE;
MotorReverse := FALSE;
CompletionLight := FALSE;

IF NOT Mode THEN
    State := IDLE;
    CompletionLatched := FALSE;

    IF ForwardButton AND NOT ReverseButton THEN
        MotorForward := TRUE;
    ELSIF ReverseButton AND NOT ForwardButton THEN
        MotorReverse := TRUE;
    END_IF;
ELSE
    CASE State OF
        IDLE:
            IF SensorA AND ButtonA THEN
                State := MOVING_TO_B;
            ELSIF SensorB THEN
                State := WAIT_B;
            ELSIF SensorC THEN
                State := WAIT_C;
            END_IF;

        MOVING_TO_B:
            IF SensorB THEN
                State := WAIT_B;
            END_IF;

        WAIT_B:
            IF NOT SensorB THEN
                State := IDLE;
            ELSIF ButtonB THEN
                State := MOVING_TO_C;
            END_IF;

        MOVING_TO_C:
            IF SensorC THEN
                State := WAIT_C;
            END_IF;

        WAIT_C:
            IF SensorC AND ButtonC THEN
                CompletionLatched := TRUE;
            END_IF;

            IF NOT SensorC THEN
                State := IDLE;
                CompletionLatched := FALSE;
            END_IF;
    END_CASE;

    MotorForward := (State = MOVING_TO_B) OR (State = MOVING_TO_C);
    CompletionLight := CompletionLatched AND SensorC;
END_IF;
END_FUNCTION_BLOCK

(* ---- public-medium-05.candidate_02.st ---- *)
TYPE AutoState : (IDLE, MOVING_TO_B, WAIT_B, MOVING_TO_C, WAIT_C);
END_TYPE;

FUNCTION_BLOCK ProductionLineControl
VAR_INPUT
    Mode : BOOL;
    ForwardButton : BOOL;
    ReverseButton : BOOL;
    SensorA : BOOL;
    SensorB : BOOL;
    SensorC : BOOL;
    ButtonA : BOOL;
    ButtonB : BOOL;
    ButtonC : BOOL;
END_VAR
VAR_OUTPUT
    MotorForward : BOOL;
    MotorReverse : BOOL;
    CompletionLight : BOOL;
END_VAR
VAR
    State : AutoState := IDLE;
    CompletionLatched : BOOL := FALSE;
END_VAR

MotorForward := FALSE;
MotorReverse := FALSE;
CompletionLight := FALSE;

IF NOT Mode THEN
    State := IDLE;
    CompletionLatched := FALSE;

    IF ForwardButton AND NOT ReverseButton THEN
        MotorForward := TRUE;
    ELSIF ReverseButton AND NOT ForwardButton THEN
        MotorReverse := TRUE;
    END_IF;
ELSE
    CASE State OF
        IDLE:
            IF SensorA AND ButtonA THEN
                State := MOVING_TO_B;
            ELSIF SensorB THEN
                State := WAIT_B;
            ELSIF SensorC THEN
                State := WAIT_C;
            END_IF;

        MOVING_TO_B:
            IF SensorB THEN
                State := WAIT_B;
            END_IF;

        WAIT_B:
            IF SensorB AND ButtonB THEN
                State := MOVING_TO_C;
            END_IF;

        MOVING_TO_C:
            IF SensorC THEN
                State := WAIT_C;
            END_IF;

        WAIT_C:
            IF SensorC AND ButtonC THEN
                CompletionLatched := TRUE;
            END_IF;

            IF NOT SensorC THEN
                State := IDLE;
                CompletionLatched := FALSE;
            END_IF;
    END_CASE;

    MotorForward := (State = MOVING_TO_B) OR (State = MOVING_TO_C);
    CompletionLight := CompletionLatched AND SensorC;
END_IF;
END_FUNCTION_BLOCK

(* ---- public-medium-05.raw_candidate_01.st ---- *)
TYPE AutoState : (IDLE, MOVING_TO_B, WAIT_B, MOVING_TO_C, WAIT_C);
END_TYPE;

FUNCTION_BLOCK ProductionLineControl
VAR_INPUT
    Mode : BOOL;
    ForwardButton : BOOL;
    ReverseButton : BOOL;
    SensorA : BOOL;
    SensorB : BOOL;
    SensorC : BOOL;
    ButtonA : BOOL;
    ButtonB : BOOL;
    ButtonC : BOOL;
END_VAR
VAR_OUTPUT
    MotorForward : BOOL;
    MotorReverse : BOOL;
    CompletionLight : BOOL;
END_VAR
VAR
    State : AutoState := IDLE;
    CompletionLatched : BOOL := FALSE;
END_VAR

MotorForward := FALSE;
MotorReverse := FALSE;
CompletionLight := FALSE;

IF NOT Mode THEN
    State := IDLE;
    CompletionLatched := FALSE;

    IF ForwardButton AND NOT ReverseButton THEN
        MotorForward := TRUE;
    ELSIF ReverseButton AND NOT ForwardButton THEN
        MotorReverse := TRUE;
    END_IF;
ELSE
    CASE State OF
        IDLE:
            IF SensorA AND ButtonA THEN
                State := MOVING_TO_B;
            ELSIF SensorB THEN
                State := WAIT_B;
            ELSIF SensorC THEN
                State := WAIT_C;
            END_IF;

        MOVING_TO_B:
            IF SensorB THEN
                State := WAIT_B;
            END_IF;

        WAIT_B:
            IF NOT SensorB THEN
                State := IDLE;
            ELSIF ButtonB THEN
                State := MOVING_TO_C;
            END_IF;

        MOVING_TO_C:
            IF SensorC THEN
                State := WAIT_C;
            END_IF;

        WAIT_C:
            IF SensorC AND ButtonC THEN
                CompletionLatched := TRUE;
            END_IF;

            IF NOT SensorC THEN
                State := IDLE;
                CompletionLatched := FALSE;
            END_IF;
    END_CASE;

    MotorForward := (State = MOVING_TO_B) OR (State = MOVING_TO_C);
    CompletionLight := CompletionLatched AND SensorC;
END_IF;
END_FUNCTION_BLOCK

(* ---- public-medium-05.raw_candidate_02.st ---- *)
TYPE AutoState : (IDLE, MOVING_TO_B, WAIT_B, MOVING_TO_C, WAIT_C);
END_TYPE;

FUNCTION_BLOCK ProductionLineControl
VAR_INPUT
    Mode : BOOL;
    ForwardButton : BOOL;
    ReverseButton : BOOL;
    SensorA : BOOL;
    SensorB : BOOL;
    SensorC : BOOL;
    ButtonA : BOOL;
    ButtonB : BOOL;
    ButtonC : BOOL;
END_VAR
VAR_OUTPUT
    MotorForward : BOOL;
    MotorReverse : BOOL;
    CompletionLight : BOOL;
END_VAR
VAR
    State : AutoState := IDLE;
    CompletionLatched : BOOL := FALSE;
END_VAR

MotorForward := FALSE;
MotorReverse := FALSE;
CompletionLight := FALSE;

IF NOT Mode THEN
    State := IDLE;
    CompletionLatched := FALSE;

    IF ForwardButton AND NOT ReverseButton THEN
        MotorForward := TRUE;
    ELSIF ReverseButton AND NOT ForwardButton THEN
        MotorReverse := TRUE;
    END_IF;
ELSE
    CASE State OF
        IDLE:
            IF SensorA AND ButtonA THEN
                State := MOVING_TO_B;
            ELSIF SensorB THEN
                State := WAIT_B;
            ELSIF SensorC THEN
                State := WAIT_C;
            END_IF;

        MOVING_TO_B:
            IF SensorB THEN
                State := WAIT_B;
            END_IF;

        WAIT_B:
            IF SensorB AND ButtonB THEN
                State := MOVING_TO_C;
            END_IF;

        MOVING_TO_C:
            IF SensorC THEN
                State := WAIT_C;
            END_IF;

        WAIT_C:
            IF SensorC AND ButtonC THEN
                CompletionLatched := TRUE;
            END_IF;

            IF NOT SensorC THEN
                State := IDLE;
                CompletionLatched := FALSE;
            END_IF;
    END_CASE;

    MotorForward := (State = MOVING_TO_B) OR (State = MOVING_TO_C);
    CompletionLight := CompletionLatched AND SensorC;
END_IF;
END_FUNCTION_BLOCK

(* ---- public-medium-06.candidate_01.st ---- *)
FUNCTION_BLOCK SlabThicknessAlarm
VAR_INPUT
    THICKNESS_FAULT : BOOL;
    THICKNESS_SIGNAL_VALID : BOOL;
    CUTTING_RUN : BOOL;
    FaultTimestamp : DINT;
    CycleTime : TIME;
END_VAR
VAR_OUTPUT
    THICKNESS_ALARM : BOOL := FALSE;
    Slab_Fault_Counter : UINT := 0;
    Slab_Runtime_Accumulator : LTIME := LTIME#0S;
    Slab_Fault_History : ARRAY[0..4] OF DINT := [0,0,0,0,0];
END_VAR
VAR
    lastValidFault : BOOL := FALSE;
    holdTimer : TIME := T#0MS;
    currentValidFault : BOOL;
    dt : LTIME;
    i : INT;
END_VAR

currentValidFault := THICKNESS_SIGNAL_VALID AND THICKNESS_FAULT;

IF NOT THICKNESS_SIGNAL_VALID THEN
    THICKNESS_ALARM := FALSE;
    holdTimer := T#0MS;
ELSE
    dt := TIME_TO_LTIME(CycleTime);

    IF currentValidFault AND NOT lastValidFault THEN
        Slab_Fault_Counter := Slab_Fault_Counter + UINT#1;

        FOR i := 4 TO 1 BY -1 DO
            Slab_Fault_History[i] := Slab_Fault_History[i - 1];
        END_FOR;

        Slab_Fault_History[0] := FaultTimestamp;
        holdTimer := T#500MS;
    END_IF;

    IF holdTimer > T#0MS THEN
        IF holdTimer > CycleTime THEN
            holdTimer := holdTimer - CycleTime;
        ELSE
            holdTimer := T#0MS;
        END_IF;
    END_IF;

    IF THICKNESS_FAULT OR (holdTimer > T#0MS) THEN
        THICKNESS_ALARM := TRUE;
    ELSE
        THICKNESS_ALARM := FALSE;
    END_IF;

    IF CUTTING_RUN AND NOT THICKNESS_FAULT THEN
        Slab_Runtime_Accumulator := Slab_Runtime_Accumulator + dt;
    END_IF;
END_IF;

lastValidFault := currentValidFault;

END_FUNCTION_BLOCK

(* ---- public-medium-06.candidate_02.st ---- *)
FUNCTION_BLOCK SlabThicknessAlarm
VAR_INPUT
    THICKNESS_FAULT : BOOL;
    THICKNESS_SIGNAL_VALID : BOOL;
    CUTTING_RUN : BOOL;
    FaultTimestamp : DINT;
    CycleTime : TIME;
END_VAR
VAR_OUTPUT
    THICKNESS_ALARM : BOOL := FALSE;
    Slab_Fault_Counter : UINT := 0;
    Slab_Runtime_Accumulator : LTIME;
    Slab_Fault_History : ARRAY[0..4] OF DINT;
END_VAR
VAR
    lastValidFault : BOOL := FALSE;
    holdTimer : TIME := T#0MS;
    initDone : BOOL := FALSE;
    i : INT;
END_VAR

// Power‑up initialisation: zero all outputs and clear holding state
IF NOT initDone THEN
    THICKNESS_ALARM := FALSE;
    Slab_Fault_Counter := 0;
    Slab_Runtime_Accumulator := LTIME#0S;
    FOR i := 0 TO 4 DO
        Slab_Fault_History[i] := 0;
    END_FOR;
    lastValidFault := FALSE;
    holdTimer := T#0MS;
    initDone := TRUE;
END_IF;

// Handle invalid signal: alarm off, no accumulation or logging
IF NOT THICKNESS_SIGNAL_VALID THEN
    THICKNESS_ALARM := FALSE;
    holdTimer := T#0MS;
    lastValidFault := FALSE;
ELSE
    // Valid signal path
    // Detect rising edge of valid fault
    IF THICKNESS_FAULT AND NOT lastValidFault THEN
        Slab_Fault_Counter := Slab_Fault_Counter + UINT#1;
        // Shift history
        FOR i := 4 TO 1 BY -1 DO
            Slab_Fault_History[i] := Slab_Fault_History[i - 1];
        END_FOR;
        Slab_Fault_History[0] := FaultTimestamp;
        holdTimer := T#500MS;
    END_IF;

    // Decrement hold timer
    IF holdTimer > T#0MS THEN
        IF holdTimer >= CycleTime THEN
            holdTimer := holdTimer - CycleTime;
        ELSE
            holdTimer := T#0MS;
        END_IF;
    END_IF;

    // Alarm condition: fault active or hold timer running
    IF THICKNESS_FAULT OR (holdTimer > T#0MS) THEN
        THICKNESS_ALARM := TRUE;
    ELSE
        THICKNESS_ALARM := FALSE;
    END_IF;

    // Accumulate runtime only when cutting, signal valid, no fault
    IF CUTTING_RUN AND NOT THICKNESS_FAULT THEN
        Slab_Runtime_Accumulator := Slab_Runtime_Accumulator + TIME_TO_LTIME(CycleTime);
    END_IF;

    // Update last valid fault state for next scan
    lastValidFault := THICKNESS_FAULT;
END_IF;

END_FUNCTION_BLOCK

(* ---- public-medium-06.raw_candidate_01.st ---- *)
FUNCTION_BLOCK SlabThicknessAlarm
VAR_INPUT
    THICKNESS_FAULT : BOOL;
    THICKNESS_SIGNAL_VALID : BOOL;
    CUTTING_RUN : BOOL;
    FaultTimestamp : DINT;
    CycleTime : TIME;
END_VAR
VAR_OUTPUT
    THICKNESS_ALARM : BOOL := FALSE;
    Slab_Fault_Counter : UINT := 0;
    Slab_Runtime_Accumulator : LTIME := LTIME#0S;
    Slab_Fault_History : ARRAY[0..4] OF DINT := [0,0,0,0,0];
END_VAR
VAR
    lastValidFault : BOOL := FALSE;
    holdTimer : TIME := T#0MS;
    currentValidFault : BOOL;
    dt : LTIME;
    i : INT;
END_VAR

currentValidFault := THICKNESS_SIGNAL_VALID AND THICKNESS_FAULT;

IF NOT THICKNESS_SIGNAL_VALID THEN
    THICKNESS_ALARM := FALSE;
    holdTimer := T#0MS;
ELSE
    dt := TIME_TO_LTIME(CycleTime);

    IF currentValidFault AND NOT lastValidFault THEN
        Slab_Fault_Counter := Slab_Fault_Counter + UINT#1;

        FOR i := 4 TO 1 BY -1 DO
            Slab_Fault_History[i] := Slab_Fault_History[i - 1];
        END_FOR;

        Slab_Fault_History[0] := FaultTimestamp;
        holdTimer := T#500MS;
    END_IF;

    IF holdTimer > T#0MS THEN
        IF holdTimer > CycleTime THEN
            holdTimer := holdTimer - CycleTime;
        ELSE
            holdTimer := T#0MS;
        END_IF;
    END_IF;

    IF THICKNESS_FAULT OR (holdTimer > T#0MS) THEN
        THICKNESS_ALARM := TRUE;
    ELSE
        THICKNESS_ALARM := FALSE;
    END_IF;

    IF CUTTING_RUN AND NOT THICKNESS_FAULT THEN
        Slab_Runtime_Accumulator := Slab_Runtime_Accumulator + dt;
    END_IF;
END_IF;

lastValidFault := currentValidFault;

END_FUNCTION_BLOCK

(* ---- public-medium-06.raw_candidate_02.st ---- *)
FUNCTION_BLOCK SlabThicknessAlarm
VAR_INPUT
    THICKNESS_FAULT : BOOL;
    THICKNESS_SIGNAL_VALID : BOOL;
    CUTTING_RUN : BOOL;
    FaultTimestamp : DINT;
    CycleTime : TIME;
END_VAR
VAR_OUTPUT
    THICKNESS_ALARM : BOOL := FALSE;
    Slab_Fault_Counter : UINT := 0;
    Slab_Runtime_Accumulator : LTIME;
    Slab_Fault_History : ARRAY[0..4] OF DINT;
END_VAR
VAR
    lastValidFault : BOOL := FALSE;
    holdTimer : TIME := T#0MS;
    initDone : BOOL := FALSE;
    i : INT;
END_VAR

// Power‑up initialisation: zero all outputs and clear holding state
IF NOT initDone THEN
    THICKNESS_ALARM := FALSE;
    Slab_Fault_Counter := 0;
    Slab_Runtime_Accumulator := LTIME#0S;
    FOR i := 0 TO 4 DO
        Slab_Fault_History[i] := 0;
    END_FOR;
    lastValidFault := FALSE;
    holdTimer := T#0MS;
    initDone := TRUE;
END_IF;

// Handle invalid signal: alarm off, no accumulation or logging
IF NOT THICKNESS_SIGNAL_VALID THEN
    THICKNESS_ALARM := FALSE;
    holdTimer := T#0MS;
    lastValidFault := FALSE;
ELSE
    // Valid signal path
    // Detect rising edge of valid fault
    IF THICKNESS_FAULT AND NOT lastValidFault THEN
        Slab_Fault_Counter := Slab_Fault_Counter + UINT#1;
        // Shift history
        FOR i := 4 TO 1 BY -1 DO
            Slab_Fault_History[i] := Slab_Fault_History[i - 1];
        END_FOR;
        Slab_Fault_History[0] := FaultTimestamp;
        holdTimer := T#500MS;
    END_IF;

    // Decrement hold timer
    IF holdTimer > T#0MS THEN
        IF holdTimer >= CycleTime THEN
            holdTimer := holdTimer - CycleTime;
        ELSE
            holdTimer := T#0MS;
        END_IF;
    END_IF;

    // Alarm condition: fault active or hold timer running
    IF THICKNESS_FAULT OR (holdTimer > T#0MS) THEN
        THICKNESS_ALARM := TRUE;
    ELSE
        THICKNESS_ALARM := FALSE;
    END_IF;

    // Accumulate runtime only when cutting, signal valid, no fault
    IF CUTTING_RUN AND NOT THICKNESS_FAULT THEN
        Slab_Runtime_Accumulator := Slab_Runtime_Accumulator + TIME_TO_LTIME(CycleTime);
    END_IF;

    // Update last valid fault state for next scan
    lastValidFault := THICKNESS_FAULT;
END_IF;

END_FUNCTION_BLOCK

(* ---- public-medium-07.candidate_01.st ---- *)
FUNCTION_BLOCK OfficeHVACControl
VAR_INPUT
    OCCUPANCY_DETECTED : BOOL;
    ENERGY_SAVING_MODE : BOOL;
    HVAC_MODE_SELECTOR : INT;
END_VAR
VAR_OUTPUT
    SUPPLY_FAN_RUN : BOOL;
    TEMP_SETPOINT_ADJUST : INT;
END_VAR
VAR
    fanDelay : TON;
    startFanCondition : BOOL;
    adjustment : INT;
END_VAR

    SUPPLY_FAN_RUN := FALSE;
    TEMP_SETPOINT_ADJUST := 0;

    startFanCondition := OCCUPANCY_DETECTED AND (HVAC_MODE_SELECTOR <> 3);
    fanDelay(IN := startFanCondition, PT := T#30S);
    SUPPLY_FAN_RUN := fanDelay.Q;

    IF HVAC_MODE_SELECTOR = 0 THEN
        IF OCCUPANCY_DETECTED THEN
            adjustment := 0;
        ELSE
            IF ENERGY_SAVING_MODE THEN
                adjustment := 3;
            ELSE
                adjustment := 2;
            END_IF;
        END_IF;
    ELSIF HVAC_MODE_SELECTOR = 1 THEN
        IF OCCUPANCY_DETECTED THEN
            adjustment := 0;
        ELSE
            adjustment := 1;
        END_IF;
    ELSIF HVAC_MODE_SELECTOR = 2 THEN
        IF OCCUPANCY_DETECTED THEN
            adjustment := 0;
        ELSE
            adjustment := 4;
        END_IF;
    ELSIF HVAC_MODE_SELECTOR = 3 THEN
        adjustment := 4;
    ELSE
        adjustment := 0;
    END_IF;

    IF adjustment > 4 THEN
        adjustment := 4;
    ELSIF adjustment < -4 THEN
        adjustment := -4;
    END_IF;

    TEMP_SETPOINT_ADJUST := adjustment;

END_FUNCTION_BLOCK

(* ---- public-medium-07.raw_candidate_01.st ---- *)
FUNCTION_BLOCK OfficeHVACControl
VAR_INPUT
    OCCUPANCY_DETECTED : BOOL;
    ENERGY_SAVING_MODE : BOOL;
    HVAC_MODE_SELECTOR : INT;
END_VAR
VAR_OUTPUT
    SUPPLY_FAN_RUN : BOOL;
    TEMP_SETPOINT_ADJUST : INT;
END_VAR
VAR
    fanDelay : TON;
    startFanCondition : BOOL;
    adjustment : INT;
END_VAR

    SUPPLY_FAN_RUN := FALSE;
    TEMP_SETPOINT_ADJUST := 0;

    startFanCondition := OCCUPANCY_DETECTED AND (HVAC_MODE_SELECTOR <> 3);
    fanDelay(IN := startFanCondition, PT := T#30S);
    SUPPLY_FAN_RUN := fanDelay.Q;

    IF HVAC_MODE_SELECTOR = 0 THEN
        IF OCCUPANCY_DETECTED THEN
            adjustment := 0;
        ELSE
            IF ENERGY_SAVING_MODE THEN
                adjustment := 3;
            ELSE
                adjustment := 2;
            END_IF;
        END_IF;
    ELSIF HVAC_MODE_SELECTOR = 1 THEN
        IF OCCUPANCY_DETECTED THEN
            adjustment := 0;
        ELSE
            adjustment := 1;
        END_IF;
    ELSIF HVAC_MODE_SELECTOR = 2 THEN
        IF OCCUPANCY_DETECTED THEN
            adjustment := 0;
        ELSE
            adjustment := 4;
        END_IF;
    ELSIF HVAC_MODE_SELECTOR = 3 THEN
        adjustment := 4;
    ELSE
        adjustment := 0;
    END_IF;

    IF adjustment > 4 THEN
        adjustment := 4;
    ELSIF adjustment < -4 THEN
        adjustment := -4;
    END_IF;

    TEMP_SETPOINT_ADJUST := adjustment;

END_FUNCTION_BLOCK

(* ---- public-medium-08.candidate_01.st ---- *)
```st
FUNCTION_BLOCK FB_IPv4Parser
VAR_INPUT
    ipText : STRING(254);
END_VAR
VAR_OUTPUT
    ipValue : UDINT;
END_VAR
VAR
    i : INT;
    len : INT;
    ch : BYTE;
    digitsInSeg : INT;
    segCount : INT;
    curVal : UDINT;
    result : UDINT;
END_VAR

ipValue := 0;
digitsInSeg := 0;
segCount := 0;
curVal := 0;
result := 0;

len := LEN(ipText);

FOR i := 1 TO len DO
    ch := ipText[i];
    IF (ch >= BYTE#48) AND (ch <= BYTE#57) THEN
        curVal := (curVal * UDINT#10) +

(* ---- public-medium-08.candidate_02.st ---- *)
FUNCTION_BLOCK FB_IPv4Parser
VAR_INPUT
    ipText : STRING(254);
END_VAR
VAR_OUTPUT
    ipValue : UDINT;
END_VAR
VAR
    i : INT;
    len : INT;
    octets : ARRAY[1..4] OF UDINT;
    curVal : UDINT;
    digitCount : INT;
    segIndex : INT;
    invalid : BOOL;
    ch : BYTE;
    digit : UDINT;
END_VAR

ipValue := 0;
invalid := FALSE;
segIndex := 1;
curVal := 0;
digitCount := 0;

FOR i := 1 TO 4 DO
    octets[i] := 0;
END_FOR;

len := LEN(ipText);

FOR i := 1 TO len DO
    ch := ipText[i];
    IF (ch >= BYTE#48) AND (ch <= BYTE#57) THEN
        digit := ch - BYTE#48;
        IF NOT invalid THEN
            IF (curVal * 10 + digit) <= 255 THEN
                curVal := curVal * 10 + digit;
                digitCount := digitCount + 1;
            ELSE
                invalid := TRUE;
            END_IF;
        END_IF;
    ELSIF ch = BYTE#46 THEN
        IF NOT invalid THEN
            IF (digitCount > 0) AND (segIndex <= 4) THEN
                octets[segIndex] := curVal;
                segIndex := segIndex + 1;
                curVal := 0;
                digitCount := 0;
            ELSE
                invalid := TRUE;
            END_IF;
        END_IF;
    ELSE
        invalid := TRUE;
    END_IF;
END_FOR;

IF NOT invalid THEN
    IF (digitCount > 0) AND (segIndex <= 4) THEN
        octets[segIndex] := curVal;
        segIndex := segIndex + 1;
    ELSIF (digitCount > 0) AND (segIndex > 4) THEN
        invalid := TRUE;
    ELSIF (digitCount = 0) THEN
        invalid := TRUE;
    END_IF;
END_IF;

IF (NOT invalid) AND (segIndex = 5) THEN
    ipValue := (octets[1] * 16777216) + (octets[2] * 65536) + (octets[3] * 256) + octets[4];
END_IF;

END_FUNCTION_BLOCK

(* ---- public-medium-08.raw_candidate_01.st ---- *)
```st
FUNCTION_BLOCK FB_IPv4Parser
VAR_INPUT
    ipText : STRING(254);
END_VAR
VAR_OUTPUT
    ipValue : UDINT;
END_VAR
VAR
    i : INT;
    len : INT;
    ch : BYTE;
    digitsInSeg : INT;
    segCount : INT;
    curVal : UDINT;
    result : UDINT;
END_VAR

ipValue := 0;
digitsInSeg := 0;
segCount := 0;
curVal := 0;
result := 0;

len := LEN(ipText);

FOR i := 1 TO len DO
    ch := ipText[i];
    IF (ch >= BYTE#48) AND (ch <= BYTE#57) THEN
        curVal := (curVal * UDINT#10) +

(* ---- public-medium-08.raw_candidate_02.st ---- *)
FUNCTION_BLOCK FB_IPv4Parser
VAR_INPUT
    ipText : STRING(254);
END_VAR
VAR_OUTPUT
    ipValue : UDINT;
END_VAR
VAR
    i : INT;
    len : INT;
    octets : ARRAY[1..4] OF UDINT;
    curVal : UDINT;
    digitCount : INT;
    segIndex : INT;
    invalid : BOOL;
    ch : BYTE;
    digit : UDINT;
END_VAR

ipValue := 0;
invalid := FALSE;
segIndex := 1;
curVal := 0;
digitCount := 0;

FOR i := 1 TO 4 DO
    octets[i] := 0;
END_FOR;

len := LEN(ipText);

FOR i := 1 TO len DO
    ch := ipText[i];
    IF (ch >= BYTE#48) AND (ch <= BYTE#57) THEN
        digit := ch - BYTE#48;
        IF NOT invalid THEN
            IF (curVal * 10 + digit) <= 255 THEN
                curVal := curVal * 10 + digit;
                digitCount := digitCount + 1;
            ELSE
                invalid := TRUE;
            END_IF;
        END_IF;
    ELSIF ch = BYTE#46 THEN
        IF NOT invalid THEN
            IF (digitCount > 0) AND (segIndex <= 4) THEN
                octets[segIndex] := curVal;
                segIndex := segIndex + 1;
                curVal := 0;
                digitCount := 0;
            ELSE
                invalid := TRUE;
            END_IF;
        END_IF;
    ELSE
        invalid := TRUE;
    END_IF;
END_FOR;

IF NOT invalid THEN
    IF (digitCount > 0) AND (segIndex <= 4) THEN
        octets[segIndex] := curVal;
        segIndex := segIndex + 1;
    ELSIF (digitCount > 0) AND (segIndex > 4) THEN
        invalid := TRUE;
    ELSIF (digitCount = 0) THEN
        invalid := TRUE;
    END_IF;
END_IF;

IF (NOT invalid) AND (segIndex = 5) THEN
    ipValue := (octets[1] * 16777216) + (octets[2] * 65536) + (octets[3] * 256) + octets[4];
END_IF;

END_FUNCTION_BLOCK

(* ---- self-easy-01.candidate_01.st ---- *)
FUNCTION_BLOCK FB
VAR_INPUT
    enable : BOOL;
    values : ARRAY[1..8] OF INT;
    count : INT;
    avgEnable : BOOL;
END_VAR
VAR_OUTPUT
    avgOut : REAL;
END_VAR
VAR
    effectiveCount : INT;
    sum : DINT;
    i : INT;
    lastAvg : REAL;
END_VAR

IF enable AND avgEnable THEN
    IF count <= 0 THEN
        avgOut := lastAvg;
    ELSE
        effectiveCount := count;
        IF effectiveCount > 8 THEN
            effectiveCount := 8;
        END_IF;
        sum := 0;
        FOR i := 1 TO effectiveCount DO
            sum := sum + INT_TO_DINT(values[i]);
        END_FOR;
        lastAvg := DINT_TO_REAL(sum) / INT_TO_REAL(effectiveCount);
        avgOut := lastAvg;
    END_IF;
ELSE
    avgOut := lastAvg;
END_IF;

END_FUNCTION_BLOCK

(* ---- self-easy-01.raw_candidate_01.st ---- *)
FUNCTION_BLOCK FB
VAR_INPUT
    enable : BOOL;
    values : ARRAY[1..8] OF INT;
    count : INT;
    avgEnable : BOOL;
END_VAR
VAR_OUTPUT
    avgOut : REAL;
END_VAR
VAR
    effectiveCount : INT;
    sum : DINT;
    i : INT;
    lastAvg : REAL;
END_VAR

IF enable AND avgEnable THEN
    IF count <= 0 THEN
        avgOut := lastAvg;
    ELSE
        effectiveCount := count;
        IF effectiveCount > 8 THEN
            effectiveCount := 8;
        END_IF;
        sum := 0;
        FOR i := 1 TO effectiveCount DO
            sum := sum + INT_TO_DINT(values[i]);
        END_FOR;
        lastAvg := DINT_TO_REAL(sum) / INT_TO_REAL(effectiveCount);
        avgOut := lastAvg;
    END_IF;
ELSE
    avgOut := lastAvg;
END_IF;

END_FUNCTION_BLOCK

(* ---- self-easy-02.candidate_01.st ---- *)
FUNCTION_BLOCK FB
VAR_INPUT
    tankLevel : REAL;
    outletFlow : REAL;
    inletPermit : BOOL;
    resetBtn : BOOL;
END_VAR
VAR_OUTPUT
    pumpRun : BOOL;
    alarmHigh : BOOL;
    alarmLow : BOOL;
    outletValveOpen : BOOL;
END_VAR
VAR
    prevResetBtn : BOOL := FALSE;
    alarmHighState : BOOL := FALSE;
    alarmLowState : BOOL := FALSE;
    resetRising : BOOL;
END_VAR

// 上升沿检测：复位按钮从 FALSE 变为 TRUE 的当拍有效
resetRising := resetBtn AND NOT prevResetBtn;

// 报警锁存，危险条件优先，复位上升沿只能清除已脱离危险的报警
alarmHighState := (tankLevel >= 85.0) OR (alarmHighState AND NOT resetRising);
alarmLowState  := (tankLevel <= 15.0) OR (alarmLowState AND NOT resetRising);

// 更新输出报警状态
alarmHigh := alarmHighState;
alarmLow  := alarmLowState;

// 泵运行：需进料许可且无任何报警
pumpRun := inletPermit AND NOT alarmHighState AND NOT alarmLowState;

// 出口阀：低报警锁存期间关闭，其他情况开启
outletValveOpen := NOT alarmLowState;

// 保存本拍按钮状态，用于下一拍上升沿判断
prevResetBtn := resetBtn;

END_FUNCTION_BLOCK

(* ---- self-easy-02.raw_candidate_01.st ---- *)
FUNCTION_BLOCK FB
VAR_INPUT
    tankLevel : REAL;
    outletFlow : REAL;
    inletPermit : BOOL;
    resetBtn : BOOL;
END_VAR
VAR_OUTPUT
    pumpRun : BOOL;
    alarmHigh : BOOL;
    alarmLow : BOOL;
    outletValveOpen : BOOL;
END_VAR
VAR
    prevResetBtn : BOOL := FALSE;
    alarmHighState : BOOL := FALSE;
    alarmLowState : BOOL := FALSE;
    resetRising : BOOL;
END_VAR

// 上升沿检测：复位按钮从 FALSE 变为 TRUE 的当拍有效
resetRising := resetBtn AND NOT prevResetBtn;

// 报警锁存，危险条件优先，复位上升沿只能清除已脱离危险的报警
alarmHighState := (tankLevel >= 85.0) OR (alarmHighState AND NOT resetRising);
alarmLowState  := (tankLevel <= 15.0) OR (alarmLowState AND NOT resetRising);

// 更新输出报警状态
alarmHigh := alarmHighState;
alarmLow  := alarmLowState;

// 泵运行：需进料许可且无任何报警
pumpRun := inletPermit AND NOT alarmHighState AND NOT alarmLowState;

// 出口阀：低报警锁存期间关闭，其他情况开启
outletValveOpen := NOT alarmLowState;

// 保存本拍按钮状态，用于下一拍上升沿判断
prevResetBtn := resetBtn;

END_FUNCTION_BLOCK

(* ---- self-hard-01.candidate_01.st ---- *)
FUNCTION_BLOCK FB
VAR_INPUT
    flowLow : BOOL;
    ackBtn : BOOL;
    sensorOK : BOOL;
END_VAR
VAR_OUTPUT
    alarmActive : BOOL;
    alarmAcked : BOOL;
    highHigh : BOOL;
END_VAR
VAR
    prevA : BOOL := FALSE;
    prevK : BOOL := FALSE;
    prevF : BOOL := FALSE;
    prevAckBtn : BOOL := FALSE;
    rising_ack : BOOL;
    A : BOOL;
    K : BOOL;
END_VAR

rising_ack := ackBtn AND NOT prevAckBtn;

A := flowLow OR (prevA AND NOT rising_ack AND NOT (prevF AND prevK));

K := A AND (NOT flowLow OR rising_ack OR (prevF AND prevA AND prevK));

alarmActive := A;
alarmAcked := K;
highHigh := NOT sensorOK;

prevA := A;
prevK := K;
prevF := flowLow;
prevAckBtn := ackBtn;

(* ---- self-hard-01.candidate_02.st ---- *)
FUNCTION_BLOCK FB
VAR_INPUT
    flowLow : BOOL;
    ackBtn : BOOL;
    sensorOK : BOOL;
END_VAR
VAR_OUTPUT
    alarmActive : BOOL;
    alarmAcked : BOOL;
    highHigh : BOOL;
END_VAR
VAR
    prevA : BOOL := FALSE;
    prevK : BOOL := FALSE;
    prevF : BOOL := FALSE;
    prevAckBtn : BOOL := FALSE;
    rising_ack : BOOL;
    A : BOOL;
    K : BOOL;
END_VAR

rising_ack := ackBtn AND NOT prevAckBtn;

A := flowLow OR (prevA AND NOT rising_ack AND NOT (prevF AND prevK));

K := A AND (NOT flowLow OR rising_ack OR (prevF AND prevA AND prevK));

alarmActive := A;
alarmAcked := K;
highHigh := NOT sensorOK;

prevA := A;
prevK := K;
prevF := flowLow;
prevAckBtn := ackBtn;

END_FUNCTION_BLOCK

(* ---- self-hard-01.raw_candidate_01.st ---- *)
FUNCTION_BLOCK FB
VAR_INPUT
    flowLow : BOOL;
    ackBtn : BOOL;
    sensorOK : BOOL;
END_VAR
VAR_OUTPUT
    alarmActive : BOOL;
    alarmAcked : BOOL;
    highHigh : BOOL;
END_VAR
VAR
    prevA : BOOL := FALSE;
    prevK : BOOL := FALSE;
    prevF : BOOL := FALSE;
    prevAckBtn : BOOL := FALSE;
    rising_ack : BOOL;
    A : BOOL;
    K : BOOL;
END_VAR

rising_ack := ackBtn AND NOT prevAckBtn;

A := flowLow OR (prevA AND NOT rising_ack AND NOT (prevF AND prevK));

K := A AND (NOT flowLow OR rising_ack OR (prevF AND prevA AND prevK));

alarmActive := A;
alarmAcked := K;
highHigh := NOT sensorOK;

prevA := A;
prevK := K;
prevF := flowLow;
prevAckBtn := ackBtn;

(* ---- self-hard-01.raw_candidate_02.st ---- *)
FUNCTION_BLOCK FB
VAR_INPUT
    flowLow : BOOL;
    ackBtn : BOOL;
    sensorOK : BOOL;
END_VAR
VAR_OUTPUT
    alarmActive : BOOL;
    alarmAcked : BOOL;
    highHigh : BOOL;
END_VAR
VAR
    prevA : BOOL := FALSE;
    prevK : BOOL := FALSE;
    prevF : BOOL := FALSE;
    prevAckBtn : BOOL := FALSE;
    rising_ack : BOOL;
    A : BOOL;
    K : BOOL;
END_VAR

rising_ack := ackBtn AND NOT prevAckBtn;

A := flowLow OR (prevA AND NOT rising_ack AND NOT (prevF AND prevK));

K := A AND (NOT flowLow OR rising_ack OR (prevF AND prevA AND prevK));

alarmActive := A;
alarmAcked := K;
highHigh := NOT sensorOK;

prevA := A;
prevK := K;
prevF := flowLow;
prevAckBtn := ackBtn;

END_FUNCTION_BLOCK

(* ---- self-hard-02.candidate_01.st ---- *)
FUNCTION_BLOCK FB
VAR_INPUT
    startBtn : BOOL;
    abortBtn : BOOL;
    setpoint : REAL;
    pv : REAL;
    maxDuration : INT;
END_VAR
VAR_OUTPUT
    elapsed : INT := 0;
    phase : INT := 0;
    timeout : BOOL := FALSE;
END_VAR
VAR
    lastStartBtn : BOOL := FALSE;
    prevPhase : INT := 0;
    prevElapsed : INT := 0;
    prevTimeout : BOOL := FALSE;
    risingStart : BOOL;
END_VAR

// 捕获上一拍输出值
prevPhase := phase;
prevElapsed := elapsed;
prevTimeout := timeout;

// 检测启动上升沿（基于上一拍 lastStartBtn）
risingStart := startBtn AND NOT lastStartBtn;

// 优先级：中止 > 新启动沿 > 运行计数/保持
IF abortBtn THEN
    // 中止：进入9，冻结计数与超时标志
    phase := 9;
    elapsed := prevElapsed;
    timeout := prevTimeout;
ELSIF risingStart THEN
    // 有效新启动：启动拍不计数
    phase := 1;
    elapsed := 0;
    timeout := FALSE;
ELSE
    // 无中止、无新启动沿
    IF (prevPhase = 1) OR (prevPhase = 2) THEN
        // 上一拍运行态，先计数一拍
        elapsed := prevElapsed + 1;

        IF elapsed >= maxDuration THEN
            // 达到超时门槛：完成态3
            timeout := TRUE;
            phase := 3;
        ELSE
            // 未超时，处理升温/保温
            timeout := FALSE;

            IF prevPhase = 1 THEN
                IF pv >= setpoint THEN
                    phase := 2; // 升温达标转保温
                ELSE
                    phase := 1; // 继续升温
                END_IF;
            ELSE
                // prevPhase = 2，保持保温
                phase := 2;
            END_IF;
        END_IF;
    ELSE
        // 上一拍非运行态（0、3、9），保持原状态
        phase := prevPhase;
        elapsed := prevElapsed;
        timeout := prevTimeout;
    END_IF;
END_IF;

// 更新上一拍启动按钮状态
lastStartBtn := startBtn;

END_FUNCTION_BLOCK

(* ---- self-hard-02.raw_candidate_01.st ---- *)
FUNCTION_BLOCK FB
VAR_INPUT
    startBtn : BOOL;
    abortBtn : BOOL;
    setpoint : REAL;
    pv : REAL;
    maxDuration : INT;
END_VAR
VAR_OUTPUT
    elapsed : INT := 0;
    phase : INT := 0;
    timeout : BOOL := FALSE;
END_VAR
VAR
    lastStartBtn : BOOL := FALSE;
    prevPhase : INT := 0;
    prevElapsed : INT := 0;
    prevTimeout : BOOL := FALSE;
    risingStart : BOOL;
END_VAR

// 捕获上一拍输出值
prevPhase := phase;
prevElapsed := elapsed;
prevTimeout := timeout;

// 检测启动上升沿（基于上一拍 lastStartBtn）
risingStart := startBtn AND NOT lastStartBtn;

// 优先级：中止 > 新启动沿 > 运行计数/保持
IF abortBtn THEN
    // 中止：进入9，冻结计数与超时标志
    phase := 9;
    elapsed := prevElapsed;
    timeout := prevTimeout;
ELSIF risingStart THEN
    // 有效新启动：启动拍不计数
    phase := 1;
    elapsed := 0;
    timeout := FALSE;
ELSE
    // 无中止、无新启动沿
    IF (prevPhase = 1) OR (prevPhase = 2) THEN
        // 上一拍运行态，先计数一拍
        elapsed := prevElapsed + 1;

        IF elapsed >= maxDuration THEN
            // 达到超时门槛：完成态3
            timeout := TRUE;
            phase := 3;
        ELSE
            // 未超时，处理升温/保温
            timeout := FALSE;

            IF prevPhase = 1 THEN
                IF pv >= setpoint THEN
                    phase := 2; // 升温达标转保温
                ELSE
                    phase := 1; // 继续升温
                END_IF;
            ELSE
                // prevPhase = 2，保持保温
                phase := 2;
            END_IF;
        END_IF;
    ELSE
        // 上一拍非运行态（0、3、9），保持原状态
        phase := prevPhase;
        elapsed := prevElapsed;
        timeout := prevTimeout;
    END_IF;
END_IF;

// 更新上一拍启动按钮状态
lastStartBtn := startBtn;

END_FUNCTION_BLOCK

(* ---- self-hard-03.candidate_01.st ---- *)
FUNCTION_BLOCK FB
VAR_INPUT
    pushEn : BOOL;
    pushItem : INT;
    popEn : BOOL;
END_VAR
VAR_IN_OUT
    fifo : ARRAY[1..8] OF INT;
END_VAR
VAR_OUTPUT
    count : INT;
    full : BOOL;
    empty : BOOL;
    head : INT;
END_VAR
VAR
    prevPush : BOOL := FALSE;
    prevPop : BOOL := FALSE;
    prevCount : INT := 0;
    oldF : ARRAY[1..8] OF INT;
    newArr : ARRAY[1..8] OF INT;
    risingPush : BOOL;
    risingPop : BOOL;
    popAct : BOOL;
    pushAct : BOOL;
    afterPopCount : INT;
    newCount : INT;
    i : INT;
END_VAR

risingPush := pushEn AND NOT prevPush;
risingPop := popEn AND NOT prevPop;

FOR i := 1 TO 8 DO
    oldF[i] := fifo[i];
END_FOR;

popAct := risingPop AND (prevCount > 0);

IF popAct THEN
    afterPopCount := prevCount - 1;
ELSE
    afterPopCount := prevCount;
END_IF;

pushAct := risingPush AND (afterPopCount < 8);

IF pushAct THEN
    newCount := afterPopCount + 1;
ELSE
    newCount := afterPopCount;
END_IF;

FOR i := 1 TO 8 DO
    newArr[i] := 0;
END_FOR;

IF popAct THEN
    IF pushAct THEN
        FOR i := 1 TO prevCount - 1 DO
            newArr[i] := oldF[i + 1];
        END_FOR;
        newArr[prevCount] := pushItem;
    ELSE
        FOR i := 1 TO prevCount - 1 DO
            newArr[i] := oldF[i + 1];
        END_FOR;
    END_IF;
ELSE
    IF pushAct THEN
        FOR i := 1 TO prevCount DO
            newArr[i] := oldF[i];
        END_FOR;
        newArr[prevCount + 1] := pushItem;
    ELSE
        FOR i := 1 TO prevCount DO
            newArr[i] := oldF[i];
        END_FOR;
    END_IF;
END_IF;

FOR i := 1 TO 8 DO
    fifo[i] := newArr[i];
END_FOR;

IF newCount > 0 THEN
    head := newArr[1];
ELSE
    head := 0;
END_IF;

count := newCount;
full := (newCount = 8);
empty := (newCount = 0);

prevPush := pushEn;
prevPop := popEn;
prevCount := newCount;
END_FUNCTION_BLOCK

(* ---- self-hard-03.raw_candidate_01.st ---- *)
FUNCTION_BLOCK FB
VAR_INPUT
    pushEn : BOOL;
    pushItem : INT;
    popEn : BOOL;
END_VAR
VAR_IN_OUT
    fifo : ARRAY[1..8] OF INT;
END_VAR
VAR_OUTPUT
    count : INT;
    full : BOOL;
    empty : BOOL;
    head : INT;
END_VAR
VAR
    prevPush : BOOL := FALSE;
    prevPop : BOOL := FALSE;
    prevCount : INT := 0;
    oldF : ARRAY[1..8] OF INT;
    newArr : ARRAY[1..8] OF INT;
    risingPush : BOOL;
    risingPop : BOOL;
    popAct : BOOL;
    pushAct : BOOL;
    afterPopCount : INT;
    newCount : INT;
    i : INT;
END_VAR

risingPush := pushEn AND NOT prevPush;
risingPop := popEn AND NOT prevPop;

FOR i := 1 TO 8 DO
    oldF[i] := fifo[i];
END_FOR

popAct := risingPop AND (prevCount > 0);

IF popAct THEN
    afterPopCount := prevCount - 1;
ELSE
    afterPopCount := prevCount;
END_IF

pushAct := risingPush AND (afterPopCount < 8);

IF pushAct THEN
    newCount := afterPopCount + 1;
ELSE
    newCount := afterPopCount;
END_IF

FOR i := 1 TO 8 DO
    newArr[i] := 0;
END_FOR

IF popAct THEN
    IF pushAct THEN
        FOR i := 1 TO prevCount - 1 DO
            newArr[i] := oldF[i + 1];
        END_FOR
        newArr[prevCount] := pushItem;
    ELSE
        FOR i := 1 TO prevCount - 1 DO
            newArr[i] := oldF[i + 1];
        END_FOR
    END_IF
ELSE
    IF pushAct THEN
        FOR i := 1 TO prevCount DO
            newArr[i] := oldF[i];
        END_FOR
        newArr[prevCount + 1] := pushItem;
    ELSE
        FOR i := 1 TO prevCount DO
            newArr[i] := oldF[i];
        END_FOR
    END_IF
END_IF

FOR i := 1 TO 8 DO
    fifo[i] := newArr[i];
END_FOR

IF newCount > 0 THEN
    head := newArr[1];
ELSE
    head := 0;
END_IF

count := newCount;
full := (newCount = 8);
empty := (newCount = 0);

prevPush := pushEn;
prevPop := popEn;
prevCount := newCount;
END_FUNCTION_BLOCK

(* ---- self-hard-04.candidate_01.st ---- *)
FUNCTION_BLOCK FB
VAR_INPUT
    demand : INT;
    runHours : ARRAY[1..5] OF LINT;
    rotated : BOOL;
END_VAR
VAR_OUTPUT
    leadPump : INT;
    lagPump : INT;
    runningCount : INT;
END_VAR
VAR
    prevLeadPump : INT := 0;
    prevLagPump : INT := 0;
    prevRunningCount : INT := 0;
    clampedDemand : INT;
    minPump : INT;
    i : INT;
END_VAR

// 裁剪需求
IF demand < 0 THEN
    clampedDemand := 0;
ELSIF demand > 5 THEN
    clampedDemand := 5;
ELSE
    clampedDemand := demand;
END_IF;

runningCount := clampedDemand;

// 计算全场最短工时泵（工时，泵号）最小
minPump := 1;
FOR i := 2 TO 5 DO
    IF (runHours[i] < runHours[minPump]) OR (runHours[i] = runHours[minPump] AND i < minPump) THEN
        minPump := i;
    END_IF;
END_FOR;

// 主泵选择
IF clampedDemand = 0 THEN
    leadPump := 0;
    lagPump := 0;
ELSE
    // 需求 > 0
    IF prevLeadPump = 0 THEN
        // 初选
        leadPump := minPump;
    ELSE
        // 已有主泵
        IF rotated AND (runHours[prevLeadPump] - runHours[minPump] > 50) THEN
            leadPump := minPump;
        ELSE
            leadPump := prevLeadPump;
        END_IF;
    END_IF;

    // 备泵选择
    IF clampedDemand < 2 THEN
        lagPump := 0;
    ELSE
        // 需求 >= 2
        IF (leadPump <> prevLeadPump) OR (clampedDemand > prevRunningCount) THEN
            // 重新选择备泵（排除当前主泵）
            lagPump := 0;
            FOR i := 1 TO 5 DO
                IF i <> leadPump THEN
                    IF lagPump = 0 THEN
                        lagPump := i;
                    ELSE
                        IF (runHours[i] < runHours[lagPump]) OR (runHours[i] = runHours[lagPump] AND i < lagPump) THEN
                            lagPump := i;
                        END_IF;
                    END_IF;
                END_IF;
            END_FOR;
        ELSE
            lagPump := prevLagPump;
        END_IF;
    END_IF;
END_IF;

// 更新上一拍状态
prevLeadPump := leadPump;
prevLagPump := lagPump;
prevRunningCount := runningCount;

END_FUNCTION_BLOCK

(* ---- self-hard-04.raw_candidate_01.st ---- *)
FUNCTION_BLOCK FB
VAR_INPUT
    demand : INT;
    runHours : ARRAY[1..5] OF LINT;
    rotated : BOOL;
END_VAR
VAR_OUTPUT
    leadPump : INT;
    lagPump : INT;
    runningCount : INT;
END_VAR
VAR
    prevLeadPump : INT := 0;
    prevLagPump : INT := 0;
    prevRunningCount : INT := 0;
    clampedDemand : INT;
    minPump : INT;
    i : INT;
END_VAR

// 裁剪需求
IF demand < 0 THEN
    clampedDemand := 0;
ELSIF demand > 5 THEN
    clampedDemand := 5;
ELSE
    clampedDemand := demand;
END_IF;

runningCount := clampedDemand;

// 计算全场最短工时泵（工时，泵号）最小
minPump := 1;
FOR i := 2 TO 5 DO
    IF (runHours[i] < runHours[minPump]) OR (runHours[i] = runHours[minPump] AND i < minPump) THEN
        minPump := i;
    END_IF;
END_FOR;

// 主泵选择
IF clampedDemand = 0 THEN
    leadPump := 0;
    lagPump := 0;
ELSE
    // 需求 > 0
    IF prevLeadPump = 0 THEN
        // 初选
        leadPump := minPump;
    ELSE
        // 已有主泵
        IF rotated AND (runHours[prevLeadPump] - runHours[minPump] > 50) THEN
            leadPump := minPump;
        ELSE
            leadPump := prevLeadPump;
        END_IF;
    END_IF;

    // 备泵选择
    IF clampedDemand < 2 THEN
        lagPump := 0;
    ELSE
        // 需求 >= 2
        IF (leadPump <> prevLeadPump) OR (clampedDemand > prevRunningCount) THEN
            // 重新选择备泵（排除当前主泵）
            lagPump := 0;
            FOR i := 1 TO 5 DO
                IF i <> leadPump THEN
                    IF lagPump = 0 THEN
                        lagPump := i;
                    ELSE
                        IF (runHours[i] < runHours[lagPump]) OR (runHours[i] = runHours[lagPump] AND i < lagPump) THEN
                            lagPump := i;
                        END_IF;
                    END_IF;
                END_IF;
            END_FOR;
        ELSE
            lagPump := prevLagPump;
        END_IF;
    END_IF;
END_IF;

// 更新上一拍状态
prevLeadPump := leadPump;
prevLagPump := lagPump;
prevRunningCount := runningCount;

END_FUNCTION_BLOCK

(* ---- self-hard-05.candidate_01.st ---- *)
FUNCTION_BLOCK FB
VAR_INPUT
    runRequest : BOOL;
    flameOK : BOOL;
    o2Valid : BOOL;
    o2PV : REAL;
    baseAir : REAL;
    resetBtn : BOOL;
END_VAR
VAR_OUTPUT
    fuelPermit : BOOL;
    trimEnable : BOOL;
    airTrim : REAL;
    airCommand : REAL;
    tripLatched : BOOL;
    o2Fault : BOOL;
END_VAR
VAR
    prevReset : BOOL;
    tripMem : BOOL;
    risingReset : BOOL;
    rawTrim : REAL;
    cmdRaw : REAL;
END_VAR

risingReset := resetBtn AND NOT prevReset;

IF (runRequest AND NOT flameOK) OR (tripMem AND NOT (risingReset AND NOT runRequest AND NOT flameOK)) THEN
    tripLatched := TRUE;
    tripMem := TRUE;
ELSE
    tripLatched := FALSE;
    tripMem := FALSE;
END_IF;

fuelPermit := runRequest AND flameOK AND NOT tripLatched;

o2Fault := (NOT o2Valid) OR (o2PV < 0.0) OR (o2PV > 21.0);

trimEnable := fuelPermit AND NOT o2Fault;

IF NOT trimEnable THEN
    airTrim := 0.0;
ELSE
    rawTrim := 2.0 * (2.0 - o2PV);
    IF rawTrim < -10.0 THEN
        airTrim := -10.0;
    ELSIF rawTrim > 10.0 THEN
        airTrim := 10.0;
    ELSE
        airTrim := rawTrim;
    END_IF;
END_IF;

IF NOT fuelPermit THEN
    airCommand := 0.0;
ELSE
    cmdRaw := baseAir + airTrim;
    IF cmdRaw < 0.0 THEN
        airCommand := 0.0;
    ELSIF cmdRaw > 100.0 THEN
        airCommand := 100.0;
    ELSE
        airCommand := cmdRaw;
    END_IF;
END_IF;

prevReset := resetBtn;

END_FUNCTION_BLOCK

(* ---- self-hard-05.raw_candidate_01.st ---- *)
FUNCTION_BLOCK FB
VAR_INPUT
    runRequest : BOOL;
    flameOK : BOOL;
    o2Valid : BOOL;
    o2PV : REAL;
    baseAir : REAL;
    resetBtn : BOOL;
END_VAR
VAR_OUTPUT
    fuelPermit : BOOL;
    trimEnable : BOOL;
    airTrim : REAL;
    airCommand : REAL;
    tripLatched : BOOL;
    o2Fault : BOOL;
END_VAR
VAR
    prevReset : BOOL;
    tripMem : BOOL;
    risingReset : BOOL;
    rawTrim : REAL;
    cmdRaw : REAL;
END_VAR

risingReset := resetBtn AND NOT prevReset;

IF (runRequest AND NOT flameOK) OR (tripMem AND NOT (risingReset AND NOT runRequest AND NOT flameOK)) THEN
    tripLatched := TRUE;
    tripMem := TRUE;
ELSE
    tripLatched := FALSE;
    tripMem := FALSE;
END_IF;

fuelPermit := runRequest AND flameOK AND NOT tripLatched;

o2Fault := (NOT o2Valid) OR (o2PV < 0.0) OR (o2PV > 21.0);

trimEnable := fuelPermit AND NOT o2Fault;

IF NOT trimEnable THEN
    airTrim := 0.0;
ELSE
    rawTrim := 2.0 * (2.0 - o2PV);
    IF rawTrim < -10.0 THEN
        airTrim := -10.0;
    ELSIF rawTrim > 10.0 THEN
        airTrim := 10.0;
    ELSE
        airTrim := rawTrim;
    END_IF;
END_IF;

IF NOT fuelPermit THEN
    airCommand := 0.0;
ELSE
    cmdRaw := baseAir + airTrim;
    IF cmdRaw < 0.0 THEN
        airCommand := 0.0;
    ELSIF cmdRaw > 100.0 THEN
        airCommand := 100.0;
    ELSE
        airCommand := cmdRaw;
    END_IF;
END_IF;

prevReset := resetBtn;

END_FUNCTION_BLOCK

(* ---- self-hard-06.candidate_01.st ---- *)
FUNCTION_BLOCK FB
VAR_INPUT
    runRequest : BOOL;
    pressure : REAL;
    pressureValid : BOOL;
    fuelFlow : REAL;
    steamFlow : REAL;
    outletCmd : INT;
    outletFeedback : INT;
    resetBtn : BOOL;
END_VAR
VAR_OUTPUT
    tripLatched : BOOL;
    fuelPermit : BOOL;
    currentCauseMask : WORD;
    latchedCauseMask : WORD;
    diagnosticActive : BOOL;
END_VAR
VAR
    prevResetBtn : BOOL := FALSE;
    stuckCount : INT := 0;
    oldTrip : BOOL;
    oldLatched : WORD;
    resetRising : BOOL;
    legalReset : BOOL;
    tripCondition : BOOL;
    bit1 : BOOL;
    bit2 : BOOL;
END_VAR

oldTrip := tripLatched;
oldLatched := latchedCauseMask;
resetRising := resetBtn AND NOT prevResetBtn;
legalReset := resetRising AND NOT runRequest AND pressureValid AND (pressure <= 4200.0);
tripCondition := runRequest AND (NOT pressureValid OR (pressure >= 4500.0));
tripLatched := tripCondition OR (oldTrip AND NOT legalReset);

currentCauseMask := 0;

IF NOT runRequest THEN
    currentCauseMask := 0;
    stuckCount := 0;
ELSIF runRequest AND NOT pressureValid THEN
    currentCauseMask := 1;
    stuckCount := 0;
ELSIF runRequest AND pressureValid AND pressure < 4500.0 THEN
    currentCauseMask := 0;
    stuckCount := 0;
ELSE
    // runRequest AND pressureValid AND pressure >= 4500.0
    IF (outletCmd >= 50) AND (outletFeedback <= 10) THEN
        IF stuckCount < 3 THEN
            stuckCount := stuckCount + 1;
        END_IF;
    ELSE
        stuckCount := 0;
    END_IF;
    bit1 := stuckCount >= 3;
    bit2 := (fuelFlow >= 4.0) AND (steamFlow <= 10.0);
    IF bit1 AND bit2 THEN
        currentCauseMask := 6;
    ELSIF bit1 THEN
        currentCauseMask := 2;
    ELSIF bit2 THEN
        currentCauseMask := 4;
    ELSE
        currentCauseMask := 8;
    END_IF;
END_IF;

IF tripLatched THEN
    latchedCauseMask := (oldLatched OR currentCauseMask) AND WORD#16#000F;
ELSE
    latchedCauseMask := 0;
END_IF;

fuelPermit := runRequest AND NOT tripLatched;
diagnosticActive := (currentCauseMask <> 0);

prevResetBtn := resetBtn;
END_FUNCTION_BLOCK

(* ---- self-hard-06.raw_candidate_01.st ---- *)
FUNCTION_BLOCK FB
VAR_INPUT
    runRequest : BOOL;
    pressure : REAL;
    pressureValid : BOOL;
    fuelFlow : REAL;
    steamFlow : REAL;
    outletCmd : INT;
    outletFeedback : INT;
    resetBtn : BOOL;
END_VAR
VAR_OUTPUT
    tripLatched : BOOL;
    fuelPermit : BOOL;
    currentCauseMask : WORD;
    latchedCauseMask : WORD;
    diagnosticActive : BOOL;
END_VAR
VAR
    prevResetBtn : BOOL := FALSE;
    stuckCount : INT := 0;
    oldTrip : BOOL;
    oldLatched : WORD;
    resetRising : BOOL;
    legalReset : BOOL;
    tripCondition : BOOL;
    bit1 : BOOL;
    bit2 : BOOL;
END_VAR

oldTrip := tripLatched;
oldLatched := latchedCauseMask;
resetRising := resetBtn AND NOT prevResetBtn;
legalReset := resetRising AND NOT runRequest AND pressureValid AND (pressure <= 4200.0);
tripCondition := runRequest AND (NOT pressureValid OR (pressure >= 4500.0));
tripLatched := tripCondition OR (oldTrip AND NOT legalReset);

currentCauseMask := 0;

IF NOT runRequest THEN
    currentCauseMask := 0;
    stuckCount := 0;
ELSIF runRequest AND NOT pressureValid THEN
    currentCauseMask := 1;
    stuckCount := 0;
ELSIF runRequest AND pressureValid AND pressure < 4500.0 THEN
    currentCauseMask := 0;
    stuckCount := 0;
ELSE
    // runRequest AND pressureValid AND pressure >= 4500.0
    IF (outletCmd >= 50) AND (outletFeedback <= 10) THEN
        IF stuckCount < 3 THEN
            stuckCount := stuckCount + 1;
        END_IF;
    ELSE
        stuckCount := 0;
    END_IF;
    bit1 := stuckCount >= 3;
    bit2 := (fuelFlow >= 4.0) AND (steamFlow <= 10.0);
    IF bit1 AND bit2 THEN
        currentCauseMask := 6;
    ELSIF bit1 THEN
        currentCauseMask := 2;
    ELSIF bit2 THEN
        currentCauseMask := 4;
    ELSE
        currentCauseMask := 8;
    END_IF;
END_IF;

IF tripLatched THEN
    latchedCauseMask := (oldLatched OR currentCauseMask) AND WORD#16#000F;
ELSE
    latchedCauseMask := 0;
END_IF;

fuelPermit := runRequest AND NOT tripLatched;
diagnosticActive := (currentCauseMask <> 0);

prevResetBtn := resetBtn;
END_FUNCTION_BLOCK

(* ---- self-hard-07.candidate_01.st ---- *)
FUNCTION_BLOCK FB
VAR_INPUT
    mode : INT;
    resetBtn : BOOL;
    scanSeconds : REAL;
    tempSP : REAL;
    tempPV : REAL;
    flowPV : REAL;
    manualFlowSP : REAL;
    manualValve : REAL;
END_VAR
VAR_OUTPUT
    flowSP : REAL;
    valveCommand : REAL;
    fault : BOOL;
    normalMode : BOOL;
END_VAR
VAR
    hasPrev : BOOL := FALSE;
    prevMode : INT := 0;
    prevReset : BOOL := FALSE;
    prevFlowSP : REAL := 0.0;
    prevValveCommand : REAL := 0.0;
    prevET : REAL := 0.0;
    prevEF : REAL := 0.0;
    resetRising : BOOL;
    eT : REAL;
    eF : REAL;
    flowRaw : REAL;
    valveRaw : REAL;
    trialT : REAL;
    trialF : REAL;
END_VAR

fault := (mode < 0) OR (mode > 2) OR (scanSeconds <= 0.0) OR (scanSeconds > 10.0);
resetRising := resetBtn AND NOT prevReset;

IF NOT hasPrev THEN
    normalMode := FALSE;
    flowSP := manualFlowSP;
    valveCommand := manualValve;
ELSIF resetRising THEN
    normalMode := FALSE;
    flowSP := manualFlowSP;
    valveCommand := manualValve;
ELSIF fault THEN
    normalMode := FALSE;
    flowSP := manualFlowSP;
    valveCommand := manualValve;
ELSIF mode <> prevMode THEN
    normalMode := FALSE;
    IF mode = 2 THEN
        flowSP := prevFlowSP;
        valveCommand := prevValveCommand;
    ELSE
        flowSP := manualFlowSP;
        valveCommand := prevValveCommand;
    END_IF;
ELSE
    normalMode := TRUE;
    IF mode = 0 THEN
        flowSP := manualFlowSP;
        valveCommand := manualValve;
    ELSIF mode = 1 THEN
        flowSP := manualFlowSP;
        eF := flowSP - flowPV;
        trialF := prevValveCommand - 2.0 * prevEF + 0.5 * eF * scanSeconds;
        valveRaw := 2.0 * eF + trialF;
        valveCommand := LIMIT(0.0, valveRaw, 100.0);
    ELSIF mode = 2 THEN
        eT := tempSP - tempPV;
        trialT := prevFlowSP - 1.0 * prevET + 0.2 * eT * scanSeconds;
        flowRaw := 1.0 * eT + trialT;
        flowSP := LIMIT(0.0, flowRaw, 50.0);
        eF := flowSP - flowPV;
        trialF := prevValveCommand - 2.0 * prevEF + 0.5 * eF * scanSeconds;
        valveRaw := 2.0 * eF + trialF;
        valveCommand := LIMIT(0.0, valveRaw, 100.0);
    END_IF;
END_IF;

prevFlowSP := flowSP;
prevValveCommand := valveCommand;
prevET := tempSP - tempPV;
prevEF := flowSP - flowPV;
prevMode := mode;
prevReset := resetBtn;
hasPrev := TRUE;

END_FUNCTION_BLOCK
